(* IEC 61131-3 sources: daoli-st-library/DL_Algo (part 6) *)

(* ---- FC_DL_HumidAirEnthalpy.st ---- *)
(*==============================================================================
 * 组件名称 (Component)  : FC_DL_HumidAirEnthalpy
 * 所属子库 (Sublibrary) : DL_Algo
 * 当前版本 (Version)    : 1.0.1
 * 组件分类 (Category)   : 函数（FUNCTION）· 湿空气热力学算法 · Level 1 算法层
 * 兼容性   (Platform)   : CODESYS 3.5 / TwinCAT 3 / 汇川 InoProShop / Schneider
 *                         Machine Expert；仅依赖 Standard.library（EXP / ABS /
 *                         MIN / MAX），零厂商方言
 * 功能描述 (Function)   : 湿空气比焓 clean-room 计算。公式链：饱和蒸汽压
 *                         p_ws 用 Magnus-Tetens（Stull 参数化，与本库
 *                         FC_DL_DewPointCalc 同系数口径 a=17.625、b=243.04，
 *                         常量复用防两套公式口径漂移）；含湿量
 *                         W = 0.622·phi·p_ws / (p - phi·p_ws)；比焓
 *                         h = 1.006·T + W·(2501 + 1.86·T)。现场用途：洁净
 *                         室/干燥房表冷器与再热功率预算、焓差控制（新风
 *                         焓 < 室内焓 才引入新风）、能耗对比。
 * 出口契约 (Exit)       : 函数返回值 = 湿空气比焓（对应规格引脚表 fEnthalpy
 *                         OUT 列），uErrorId 为 VAR_OUTPUT。异常路径返回
 *                         确定值 0.0，绝不返回未初始化值。
 * 开源溯源 (Origin)     : oscat-building / psychrolib。行为定义对标 OSCAT
 *                         Building 的 AIR_ENTHALPY（0~100 摄氏度域）与
 *                         PsychroLib GetMoistAirEnthalpy 的公开物理公式链；
 *                         公开物理公式无版权义务，不读取、不复制任何源码行，
 *                         100% clean-room 重写并按本库防御规范加严。
 * 属主转移 (R23 裁定)   : Magnus-Tetens 常数（a=17.625、b=243.04）唯一属主
 *                         自 R23 起为 FC_DL_VaporPressureSat；本件内联
 *                         DL_AIR_A / DL_AIR_B 为属主口径的历史引用，本版
 *                         仅声明、逻辑零改动，口径变更以属主件为单一事实源。
 * 规格偏离留档 (R11)    : 规格引脚表 uErrorId 原标注 0001_0203；按第 0 节
 *                         公约 0.7（优先级高于逐组件条款）沿用所在子库
 *                         DL_Algo 既有故障码段 16#0002_xxxx，细分 17xx
 *                         （15xx 露点 / 16xx 流量已占用，顺延无冲突）。
 * 验收向量 (Acceptance) :
 *   V1 T=25.0 RH=60.0 p=101.325：h 约 55.39 kJ/kg 干空气（容差 0.5）；
 *   V2 T=0.0 RH=100.0：h 约 9.44 kJ/kg 干空气（容差 0.5），uErrorId=0；
 *   V3 T=40.0 RH=1.0：干空气端下界，h 约 41.41（容差 0.5）；
 *   V4 RH=0.0：钳位至 1.0，uErrorId=16#0002_1701，照算不发散；
 *   V5 T=150.0：钳位至 100.0，uErrorId=16#0002_1701；
 *   V6 fAtmPress=200.0：钳位至 110.0，uErrorId=16#0002_1702；
 *   V7 T=100.0 RH=100.0：饱和退化分母保护，uErrorId=16#0002_1703，
 *      返回有限确定值；
 *   V8 NaN 输入：拒绝并返回 0.0，uErrorId=16#0002_0004（DL_Algo 公共码）。
 * 故障码表 (Error codes):
 *   16#0002_1701【信息级】温度/湿度越界已钳位照算 / 16#0002_1702【信息级】
 *   大气压越界已钳位照算 / 16#0002_1703【信息级】饱和退化分母已保护 /
 *   16#0002_0004【信息级】输入非有限值已拒绝。全部信息级，本函数无
 *   bError 引脚，故障分级判读经 uErrorId。
 * 修订历史 (Revision)   :
 *   2026-11-15  v1.0.0  首版入库（Round 05 · OSCAT Building 开组 · DL_Algo 补强）
 *============================================================================*)

(*-----------------------------------------------------------------------------
 * 调用示例 (Instance guide)：
 *   fHSupply := FC_DL_HumidAirEnthalpy(fTempC := stAHU.fSupplyT,
 *                                      fRelHum := stAHU.fSupplyRh,
 *                                      uErrorId => uHErr);
 *   fHOutdoor := FC_DL_HumidAirEnthalpy(fTempC := stMet.fTemp,
 *                                       fRelHum := stMet.fRh,
 *                                       fAtmPress := 100.8);
 *   焓差控制联锁：IF (fHOutdoor < fHReturn - 2.0) THEN bFreshAirOk := TRUE;
 *   仅当 uErrorId = 0 时焓值才可用于联锁判断；钳位拍（1701/1702/1703）
 *   的结果按趋势参考处理。
 *----------------------------------------------------------------------------*)

(*-----------------------------------------------------------------------------
 * 常见误用与现场提示 (Field notes)：
 *   1 输入必须是干球温度 + 相对湿度百分数；给成湿球温度或绝对湿度会得到
 *     荒谬结果。露点请先经 FC_DL_DewPointCalc 反算而不是反复试凑本函数。
 *   2 高原/密闭厂房务必传真实大气压 fAtmPress：海拔 2000m 处大气压约
 *     79.5 kPa 已低于钳位下限 80，含湿量 W 会系统性偏小，影响表冷选型。
 *   3 返回值为「每公斤干空气」比焓，做能量平衡时风量要乘干空气密度换算，
 *     勿直接乘湿空气总流量。
 *   4 100 摄氏度/100% 附近 W 发散是物理事实（水的沸点），本函数以 1 Pa
 *     分母下限保护输出有限值，但该域结果无工程意义，勿用于工艺联锁。
 *   5 纯计算无状态，可放心放入高速任务；输入应来自滤波后的温湿度信号。
 *----------------------------------------------------------------------------*)
FUNCTION FC_DL_HumidAirEnthalpy : REAL
VAR_INPUT
    fTempC    : REAL;                    // 干球温度 [摄氏度]，有效域 0.0..100.0 / Dry-bulb temperature [degC], valid range 0.0..100.0
    fRelHum   : REAL;                    // 相对湿度 [百分数]，有效域 1.0..100.0 / Relative humidity [percent], valid range 1.0..100.0
    fAtmPress : REAL := 101.325;         // 大气压 [kPa]，默认标准大气，有效域 80.0..110.0 / Atmospheric pressure [kPa], default standard atmosphere
END_VAR
VAR_OUTPUT
    uErrorId  : UDINT;                   // 故障码，16#0002_0000 = 无故障 / Error code, 16#0002_0000 = no error
END_VAR
VAR
    fTEff     : REAL;                    // 钳位后的生效温度 [摄氏度] / Effective clamped temperature [degC]
    fRhEff    : REAL;                    // 钳位后的生效湿度 [百分数] / Effective clamped humidity [percent]
    fPEff     : REAL;                    // 钳位后的生效大气压 [kPa] / Effective clamped atmospheric pressure [kPa]
    fPws      : REAL;                    // 饱和蒸汽压 [Pa] / Saturation vapor pressure [Pa]
    fPhi      : REAL;                    // 相对湿度份额 [1] / Relative humidity fraction [1]
    fPAbs     : REAL;                    // 绝对大气压 [Pa] / Absolute atmospheric pressure [Pa]
    fPv       : REAL;                    // 水汽分压 [Pa] / Water vapor partial pressure [Pa]
    fDenom    : REAL;                    // 含湿量分母 [Pa] / Humidity ratio denominator [Pa]
    fHumRatio : REAL;                    // 含湿量 [kg 水汽/kg 干空气] / Humidity ratio [kg vapor per kg dry air]
END_VAR
VAR CONSTANT
    DL_AIR_A       : REAL := 17.625;     // Magnus 系数 a [1]，与 FC_DL_DewPointCalc 同口径 / Magnus coefficient a [1], same as dew point FC
    DL_AIR_B       : REAL := 243.04;     // Magnus 系数 b [摄氏度] / Magnus coefficient b [degC]
    DL_AIR_E0      : REAL := 611.2;      // 0 摄氏度饱和水汽压 [Pa] / Saturation vapor pressure at 0 degC [Pa]
    DL_AIR_T_MIN   : REAL := 0.0;        // 温度有效域下限 [摄氏度] / Temperature valid range low [degC]
    DL_AIR_T_MAX   : REAL := 100.0;      // 温度有效域上限 [摄氏度] / Temperature valid range high [degC]
    DL_AIR_RH_MIN  : REAL := 1.0;        // 湿度钳位下限 [百分数]，防 W 比值超线性 / Humidity clamp floor [percent]
    DL_AIR_P_MIN   : REAL := 80.0;       // 大气压钳位下限 [kPa] / Pressure clamp floor [kPa]
    DL_AIR_P_MAX   : REAL := 110.0;      // 大气压钳位上限 [kPa] / Pressure clamp ceiling [kPa]
    DL_AIR_MW      : REAL := 0.622;      // 干空气/水汽摩尔比 [kg/kg] / Molar mass ratio dry air to vapor [kg/kg]
    DL_AIR_CP_DRY  : REAL := 1.006;      // 干空气比热 [kJ/(kg·K)] / Dry air specific heat [kJ/(kg*K)]
    DL_AIR_HFG0    : REAL := 2501.0;     // 0 摄氏度水汽化潜热 [kJ/kg] / Latent heat of vaporization at 0 degC [kJ/kg]
    DL_AIR_CP_VAP  : REAL := 1.86;       // 水汽比热 [kJ/(kg·K)] / Vapor specific heat [kJ/(kg*K)]
    DL_AIR_DENOM_MIN : REAL := 1.0;      // 含湿量分母保护下限 [Pa] / Humidity ratio denominator floor [Pa]
    DL_AIR_EPS     : REAL := 1.0E-6;     // 浮点判零容差 / Float zero tolerance
    DL_AIR_INF_MAX : REAL := 1.0E30;     // 有限值判定幅值上限 / Magnitude bound for finite-value check
END_VAR

(*------------------------------------------------------------------------------
 * 段 1｜出口默认值（IEC 61131-3 强制）：入口即赋确定值，任何提前 RETURN
 *      前输出已确定；异常路径返回 0.0（确定值口径）
 *      Exit defaults (mandatory): outputs assigned deterministically on entry
 *-----------------------------------------------------------------------------*)
FC_DL_HumidAirEnthalpy := 0.0;                    // 返回值（比焓）默认置零 / Return value (enthalpy) preset to zero
uErrorId := 16#0002_0000;                         // 故障码先清零 / Error code cleared first
fTEff := DL_AIR_T_MIN;                            // 温度预置域下限 / Temperature preset to domain floor
fRhEff := DL_AIR_RH_MIN;                          // 湿度预置钳位下限 / Humidity preset to clamp floor
fPEff := 101.325;                                 // 大气压预置标准值 [kPa] / Pressure preset to standard value [kPa]

(*------------------------------------------------------------------------------
 * 段 2｜非有限值防御（公约 0.8）：全部 REAL 输入（含看似常量的大气压）
 *      先做 fX <> fX 检测再比较；命中即拒绝并返回确定值
 *      Non-finite defense: all REAL inputs checked before any comparison
 *-----------------------------------------------------------------------------*)
IF (fTempC <> fTempC) OR (ABS(fTempC) > DL_AIR_INF_MAX)
   OR (fRelHum <> fRelHum) OR (ABS(fRelHum) > DL_AIR_INF_MAX)
   OR (fAtmPress <> fAtmPress) OR (ABS(fAtmPress) > DL_AIR_INF_MAX) THEN
    uErrorId := 16#0002_0004;                     // 输入非有限值已拒绝（DL_Algo 公共码）/ Non-finite input rejected
    FC_DL_HumidAirEnthalpy := 0.0;
    RETURN;
END_IF

(*------------------------------------------------------------------------------
 * 段 3｜温度钳位 [0, 100]：越界信息级码，钳位后照算（R21：不构成故障）
 *      Temperature clamping into [0, 100], info-level code, compute on
 *-----------------------------------------------------------------------------*)
IF (fTempC < DL_AIR_T_MIN) OR (fTempC > DL_AIR_T_MAX) THEN
    fTEff := MIN(MAX(fTempC, DL_AIR_T_MIN), DL_AIR_T_MAX);  // 双侧钳位到有效域 / Two-sided clamp into valid range
    uErrorId := 16#0002_1701;                     // 温度越界已钳位 / Temperature out of range clamped
ELSE
    fTEff := fTempC;                              // 合法温度原值生效 / Valid temperature applied as-is
END_IF

(*------------------------------------------------------------------------------
 * 段 4｜湿度钳位 [1, 100]（公约 0.3 限幅域一致）：下限防 W 发散，上限防
 *      超饱和非物理输入；量纲注释 [百分数] 与限幅域一致（R20）
 *      Humidity clamping into [1, 100], floor guards W divergence
 *-----------------------------------------------------------------------------*)
IF (fRelHum < DL_AIR_RH_MIN) OR (fRelHum > 100.0) THEN
    fRhEff := MIN(MAX(fRelHum, DL_AIR_RH_MIN), 100.0);      // 双侧钳位 / Two-sided clamp
    uErrorId := 16#0002_1701;                     // 湿度越界已钳位 / Humidity out of range clamped
ELSE
    fRhEff := fRelHum;                            // 合法湿度原值生效 / Valid humidity applied as-is
END_IF

(*------------------------------------------------------------------------------
 * 段 5｜大气压钳位 [80, 110] kPa：覆盖海平面 ~ 海拔 2000m 工况域
 *      Atmospheric pressure clamping into [80, 110] kPa
 *-----------------------------------------------------------------------------*)
IF (fAtmPress < DL_AIR_P_MIN) OR (fAtmPress > DL_AIR_P_MAX) THEN
    fPEff := MIN(MAX(fAtmPress, DL_AIR_P_MIN), DL_AIR_P_MAX);  // 双侧钳位 / Two-sided clamp
    uErrorId := 16#0002_1702;                     // 大气压越界已钳位 / Pressure out of range clamped
ELSE
    fPEff := fAtmPress;                           // 合法大气压原值生效 / Valid pressure applied as-is
END_IF

(*------------------------------------------------------------------------------
 * 段 6｜Magnus-Tetens 饱和蒸汽压：与 FC_DL_DewPointCalc 同系数口径，
 *      常量复用防两套公式口径漂移（热平衡算得平）
 *      Magnus-Tetens saturation vapor pressure, same coefficients as dew
 *      point FC, shared constants prevent formula drift
 *-----------------------------------------------------------------------------*)
fPws := DL_AIR_E0 * EXP(DL_AIR_A * fTEff / (DL_AIR_B + fTEff));  // 饱和蒸汽压 [Pa] / Saturation vapor pressure [Pa]

(*------------------------------------------------------------------------------
 * 段 7｜含湿量 W = 0.622·phi·p_ws / (p - phi·p_ws)：分母防除零/防退化
 *      Humidity ratio with denominator guard (divide-by-zero protected)
 *-----------------------------------------------------------------------------*)
fPhi := fRhEff / 100.0;                           // 相对湿度份额 [1] / RH fraction [1]
fPAbs := fPEff * 1000.0;                          // 大气压 kPa → Pa / Pressure kPa converted to Pa
fPv := fPhi * fPws;                               // 水汽分压 [Pa] / Vapor partial pressure [Pa]
fDenom := fPAbs - fPv;                            // 含湿量分母 [Pa] / Denominator [Pa]
IF fPAbs <= DL_AIR_EPS THEN
    uErrorId := 16#0002_1702;                     // 绝对压力退化按大气压类信息级处理 / Degenerate pressure, info code
    FC_DL_HumidAirEnthalpy := 0.0;
    RETURN;
END_IF
IF fDenom <= DL_AIR_DENOM_MIN THEN
    fPv := fPAbs - DL_AIR_DENOM_MIN;              // 饱和退化保护：水汽分压钳至分母下限之上 / Saturation degenerate guard
    uErrorId := 16#0002_1703;                     // 分母退化已保护（100 度/100% 物理发散域） / Degenerate denominator protected
END_IF
fHumRatio := DL_AIR_MW * fPv / (fPAbs - fPv);     // 含湿量 [kg 水汽/kg 干空气] / Humidity ratio [kg/kg dry air]
                                                  // 分母 = fPAbs - fPv ≥ DL_AIR_DENOM_MIN，防除零成立
(*------------------------------------------------------------------------------
 * 段 8｜比焓 h = 1.006·T + W·(2501 + 1.86·T)：显热 + 水汽潜热项
 *      Specific enthalpy: sensible dry-air term plus vapor latent term
 *-----------------------------------------------------------------------------*)
FC_DL_HumidAirEnthalpy := DL_AIR_CP_DRY * fTEff + fHumRatio * (DL_AIR_HFG0 + DL_AIR_CP_VAP * fTEff);
                                                  // 湿空气比焓 [kJ/kg 干空气] / Moist air specific enthalpy [kJ/kg dry air]
END_FUNCTION

(* ---- FC_DL_HystCounterStep.st ---- *)
(*==============================================================================
 * 名称 : FC_DL_HystCounterStep —— 迟滞跨带计数器（上穿 +1 下穿 -1，带位记忆经 nBand 回写）
 * 分类 / 前缀 / 版本 : DL_Algo / FC_DL_ / 1.0.0
 * 溯源 : 开源语义参考（OSCAT/AixOCAT 族，MIT）或 clean-room IEC 实现，未复制源码
 * 平台 : 纯 IEC 61131-3
 * 功能说明 : 以 fUpTh/fDnTh 构成上下带界、fHyst 为校验用回差参考：fIn 上穿
 *            fUpTh 计数 +1，下穿 fDnTh 计数 -1，两界之间不动作（迟滞死区）。
 *            带位记忆 nBand（-1/0/+1）经 VAR_IN_OUT 由调用方持有，保证停在
 *            界外不重复计数、须先穿越对侧门限才反向计数。计数钳位 [nMin,nMax]。
 *            边界处理：fDnTh>=fUpTh、fHyst<0、nMin>nMax 判参数非法；输入
 *            非有限（NaN/±Inf）置 eErr，两种故障下 nBand 保持原值不误动。
 * 错误码 : 16#0001_1C03 = 门限/回差/钳位区间参数非法，或输入非有限（NaN/±Inf）
 *          eErr=0 且 bValid=TRUE 表示计数结果可用（调用方须把返回值写回计数变量）
 * 状态机 : R6 标注 N/A（纯函数无顺序状态，带位记忆由调用方经 nBand 持有，以本节替代 ELSE 兜底）
 * 红线 : R1/R2/R3 ✓ 零全局/零IO/纯IEC ｜ R4 ✓ 非有限拦截/门限校验 ｜ R10 ✓ 标准转换 ｜ R11 ✓ 分号收尾 ｜ R15 ✓ 无保留字撞名
 * 修订记录 : 2026-11-23 v1.0.0 首次入库（R76）
 *============================================================================*)
FUNCTION FC_DL_HystCounterStep : INT
VAR_INPUT
    nCount : INT;      // 当前计数（调用方持有，返回值须写回）/ current count, caller-held
    fIn    : LREAL;    // 被监视输入量 [工程单位] / monitored input value
    fUpTh  : LREAL;    // 上穿计数门限 [工程单位] / up-cross counting threshold
    fDnTh  : LREAL;    // 下穿计数门限 [工程单位] / down-cross counting threshold
    fHyst  : LREAL;    // 回差参考量（须 >=0）[工程单位] / hysteresis reference, must be >= 0
    nMin   : INT;      // 计数下限 [次] / count lower clamp
    nMax   : INT;      // 计数上限 [次] / count upper clamp
END_VAR
VAR_IN_OUT
    nBand  : INT;      // 带位记忆 -1/0/+1（调用方持有回写）/ band memory, caller-held
END_VAR
VAR_OUTPUT
    eErr   : UDINT;    // 故障码，0=正常，1C03=参数非法或非有限 / error code
    bError : BOOL;     // TRUE=本件发生故障 / TRUE when fault occurred
    bValid : BOOL;     // TRUE=计数结果可用 / TRUE when count result is usable
END_VAR
VAR
    _nRet : INT;       // 计数中间值 / count intermediate
END_VAR

FC_DL_HystCounterStep := nCount;             // 返回值预设原计数 / preset return to input count
eErr   := 16#0000_0000;                      // 故障码清零 / clear error code
bError := FALSE;                             // 故障标志清零 / clear error flag
bValid := TRUE;                              // 预设输出可用 / preset valid flag

IF (fIn <> fIn) OR ((fIn - fIn) <> (fIn - fIn))          // fIn 非有限 / NaN or infinite
   OR (fUpTh <> fUpTh) OR ((fUpTh - fUpTh) <> (fUpTh - fUpTh))   // fUpTh 非有限 / NaN or infinite
   OR (fDnTh <> fDnTh) OR ((fDnTh - fDnTh) <> (fDnTh - fDnTh))   // fDnTh 非有限 / NaN or infinite
   OR (fHyst <> fHyst) OR ((fHyst - fHyst) <> (fHyst - fHyst)) THEN  // fHyst 非有限 / NaN or infinite
    eErr   := 16#0001_1C03;                  // 置非有限故障码 / set non-finite code
    bError := TRUE;                          // 置故障标志 / set error flag
    bValid := FALSE;                         // 输出不可用 / outputs not usable
    RETURN;                                  // nBand 冻结原值 / freeze band unchanged
END_IF

IF (fDnTh >= fUpTh) OR (fHyst < 0.0) OR (nMin > nMax) THEN    // 参数合法性校验 / parameter validity check
    eErr   := 16#0001_1C03;                  // 置参数非法码 / set invalid-parameter code
    bError := TRUE;                          // 置故障标志 / set error flag
    bValid := FALSE;                         // 输出不可用 / outputs not usable
    RETURN;                                  // nBand 冻结原值 / freeze band unchanged
END_IF

_nRet := nCount;                             // 取当前计数 / take current count

IF (fIn >= fUpTh) AND (nBand < 1) THEN       // 上穿且非已在高带 / up-cross and not already high
    _nRet := _nRet + 1;                      // 计数 +1 / bump count up
    nBand := 1;                              // 记忆进入高带 / memorize high band
ELSIF (fIn <= fDnTh) AND (nBand > -1) THEN   // 下穿且非已在低带 / down-cross and not already low
    _nRet := _nRet - 1;                      // 计数 -1 / bump count down
    nBand := -1;                             // 记忆进入低带 / memorize low band
ELSIF (fIn > fDnTh) AND (fIn < fUpTh) THEN   // 落入迟滞死区 / inside hysteresis deadband
    nBand := 0;                              // 记忆回到中性带 / memorize neutral band
END_IF

IF _nRet < nMin THEN                         // 计数下限钳位 / clamp lower
    _nRet := nMin;                           // 钳到下限 / clamp to lower
END_IF
IF _nRet > nMax THEN                         // 计数上限钳位 / clamp upper
    _nRet := nMax;                           // 钳到上限 / clamp to upper
END_IF

FC_DL_HystCounterStep := _nRet;              // 回写计数结果 / write back count

END_FUNCTION

(* ---- FC_DL_HystLatchAlarm.st ---- *)
(*==============================================================================
 * 名称 : FC_DL_HystLatchAlarm —— 迟滞触发 + 手动复位锁存报警（状态经 VAR_IN_OUT 由调用方持有）
 * 分类 / 前缀 / 版本 : DL_Algo / FC_DL_ / 1.0.0
 * 溯源 : 开源语义参考（OSCAT/AixOCAT 族，MIT）或 clean-room IEC 实现，未复制源码
 * 平台 : 纯 IEC 61131-3
 * 功能说明 : fIn 上穿 fOn 置位报警并锁存；降到 fOff 以下不自动清除，仅当
 *            bReset=TRUE 才复位（复位后若 fIn 仍 >= fOn 则同拍重新置位，
 *            天然防「复位即复报」盲区）。锁存状态 nState 经 VAR_IN_OUT 由
 *            调用方持有（0=正常 / 1=报警锁存），返回值 = 报警有效电平。
 *            边界处理：fOn<fOff 判参数非法（迟滞反向无意义）；输入非有限
 *            （NaN/±Inf）置 eErr，两种故障下 nState 保持原值不误动。
 * 错误码 : 16#0001_1C02 = 门限次序非法（fOn<fOff），或输入非有限（NaN/±Inf）
 *          eErr=0 且 bValid=TRUE 表示报警电平与 nState 可用
 * 状态机 : R6 标注 N/A（纯函数无顺序状态，锁存态由调用方经 nState 持有，以本节替代 ELSE 兜底）
 * 红线 : R1/R2/R3 ✓ 零全局/零IO/纯IEC ｜ R4 ✓ 非有限拦截/门限校验 ｜ R10 ✓ 标准转换 ｜ R11 ✓ 分号收尾 ｜ R15 ✓ 无保留字撞名
 * 修订记录 : 2026-11-23 v1.0.0 首次入库（R76）
 *============================================================================*)
FUNCTION FC_DL_HystLatchAlarm : BOOL
VAR_INPUT
    fIn    : LREAL;    // 被监视输入量 [工程单位] / monitored input value
    fOn    : LREAL;    // 报警置位门限 [工程单位] / alarm set threshold
    fOff   : LREAL;    // 迟滞参考门限（仅作参数校验：要求 fOn >= fOff）[工程单位] / hysteresis reference, param check only
    bReset : BOOL;     // 复位指令（沿/电平均可，调用方决定）/ reset command
END_VAR
VAR_IN_OUT
    nState : INT;      // 锁存状态 0=正常 1=报警（调用方持有回写）/ latched state, caller-held
END_VAR
VAR_OUTPUT
    eErr   : UDINT;    // 故障码，0=正常，1C02=参数非法或非有限 / error code
    bError : BOOL;     // TRUE=本件发生故障 / TRUE when fault occurred
    bValid : BOOL;     // TRUE=报警电平可用 / TRUE when alarm level is usable
END_VAR

FC_DL_HystLatchAlarm := FALSE;               // 报警电平预设 FALSE / preset alarm to FALSE
eErr   := 16#0000_0000;                      // 故障码清零 / clear error code
bError := FALSE;                             // 故障标志清零 / clear error flag
bValid := TRUE;                              // 预设输出可用 / preset valid flag

IF (fIn <> fIn) OR ((fIn - fIn) <> (fIn - fIn))          // fIn 非有限 / NaN or infinite
   OR (fOn <> fOn) OR ((fOn - fOn) <> (fOn - fOn))        // fOn 非有限 / NaN or infinite
   OR (fOff <> fOff) OR ((fOff - fOff) <> (fOff - fOff)) THEN  // fOff 非有限 / NaN or infinite
    eErr   := 16#0001_1C02;                  // 置非有限故障码 / set non-finite code
    bError := TRUE;                          // 置故障标志 / set error flag
    bValid := FALSE;                         // 输出不可用 / outputs not usable
    RETURN;                                  // nState 冻结原值，不误动 / freeze state unchanged
END_IF

IF fOn < fOff THEN                           // 迟滞反向：参数非法 / reversed hysteresis invalid
    eErr   := 16#0001_1C02;                  // 置参数非法码 / set invalid-parameter code
    bError := TRUE;                          // 置故障标志 / set error flag
    bValid := FALSE;                         // 输出不可用 / outputs not usable
    RETURN;                                  // nState 冻结原值 / freeze state unchanged
END_IF

IF bReset THEN                               // 手动复位优先（先清后判）/ reset first, judge after
    nState := 0;                             // 清除锁存 / clear latch
END_IF
IF nState = 0 THEN                           // 非锁存态才可置位 / only unlatched state can set
    IF fIn >= fOn THEN                       // 上穿置位门限 / rising past set threshold
        nState := 1;                         // 置位并锁存 / set and latch
    END_IF
END_IF

FC_DL_HystLatchAlarm := (nState = 1);        // 回写报警电平 / write back alarm level

END_FUNCTION

(* ---- FC_DL_HystTimeQualified.st ---- *)
(*==============================================================================
 * 名称 : FC_DL_HystTimeQualified —— 迟滞 + 时间确认翻转（确认计时由调用方 TON 持有）
 * 分类 / 前缀 / 版本 : DL_Algo / FC_DL_ / 1.0.0
 * 溯源 : 开源语义参考（OSCAT/AixOCAT 族，MIT）或 clean-room IEC 实现，未复制源码
 * 平台 : 纯 IEC 61131-3
 * 功能说明 : 输出翻转需时间确认：bRawIn=FALSE 时输出立即 FALSE 且确认计时
 *            清零（tNewElapsed=T#0s）；bRawIn=TRUE 且输出当前 FALSE 时，仅当
 *            调用方 TON 累计 tElapsed >= tQual 才翻转 TRUE；输出已 TRUE 且
 *            原始输入仍 TRUE 则保持。tElapsed 语义 = 调用方 TON.ET（bRawIn
 *            期间单调增长），tNewElapsed 回传给调用方供下一拍使用。
 *            边界处理：tQual<=T#0s 视为立即确认（0 时延合法用法）；
 *            bPrevOut=TRUE 而 bRawIn=FALSE 时立即翻 FALSE（OFF 无延时）。
 * 错误码 : 16#0001_1C04 为本件预留码位（当前实现无故障路径），eErr 恒 0、bValid 恒 TRUE
 * 状态机 : R6 标注 N/A（纯函数无顺序状态，确认计时由调用方 TON 持有，以本节替代 ELSE 兜底）
 * 红线 : R1/R2/R3 ✓ 零全局/零IO/纯IEC ｜ R4 ✓ 时间比较口径明确 ｜ R10 ✓ 标准转换 ｜ R11 ✓ 分号收尾 ｜ R15 ✓ 无保留字撞名
 * 修订记录 : 2026-11-23 v1.0.0 首次入库（R76）
 *============================================================================*)
FUNCTION FC_DL_HystTimeQualified : BOOL
VAR_INPUT
    bRawIn   : BOOL;   // 原始输入（未经确认）/ raw input before qualification
    tQual    : TIME;   // 确认时长门限 [ms] / qualification duration threshold
    bPrevOut : BOOL;   // 上一拍输出（调用方持有）/ previous output, caller-held
    tElapsed : TIME;   // 调用方 TON 累计确认时间 [ms] / caller-held TON elapsed time
END_VAR
VAR_OUTPUT
    tNewElapsed : TIME;    // 回传确认时间（供调用方下一拍使用）/ elapsed time passed back to caller
    eErr        : UDINT;   // 故障码，0=正常（本件无故障路径）/ error code, 0=ok (no fault path)
    bError      : BOOL;    // 故障标志，恒 FALSE / error flag, always FALSE
    bValid      : BOOL;    // TRUE=输出与计时可用，恒 TRUE / TRUE when outputs are usable
END_VAR

eErr        := 16#0000_0000;             // 故障码清零 / clear error code
bError      := FALSE;                    // 故障标志清零 / clear error flag
bValid      := TRUE;                     // 本件无故障路径，恒可用 / always valid
tNewElapsed := T#0s;                     // 确认计时预设清零 / preset elapsed to zero

IF NOT bRawIn THEN                       // 原始输入失效：OFF 无延时 / raw input low: immediate off
    FC_DL_HystTimeQualified := FALSE;    // 输出立即 FALSE / output FALSE immediately
    tNewElapsed := T#0s;                 // 确认计时清零（调用方应同步复位 TON）/ reset qualification timer
    RETURN;                              // 提前收口 / early exit
END_IF

tNewElapsed := tElapsed;                 // 原始输入有效：计时透传 / raw high: pass timer through

IF bPrevOut THEN                         // 输出已 TRUE 且原始输入仍 TRUE / already on and raw high
    FC_DL_HystTimeQualified := TRUE;     // 保持 TRUE / keep TRUE
ELSIF tElapsed >= tQual THEN             // 确认计时到限 / qualification time reached
    FC_DL_HystTimeQualified := TRUE;     // 翻转为 TRUE / flip to TRUE
ELSE                                     // 确认时间未到 / qualification not reached
    FC_DL_HystTimeQualified := FALSE;    // 维持 FALSE / keep FALSE
END_IF

END_FUNCTION

(* ---- FC_DL_HystWindow3.st ---- *)
(*==============================================================================
 * 名称 : FC_DL_HystWindow3 —— 三带迟滞带位判定（低/中/高，回差记忆由调用方持有）
 * 分类 / 前缀 / 版本 : DL_Algo / FC_DL_ / 1.0.0
 * 溯源 : 开源语义参考（OSCAT/AixOCAT 族，MIT）或 clean-room IEC 实现，未复制源码
 * 平台 : 纯 IEC 61131-3
 * 功能说明 : 返回三带带位：0=低带、1=中带、2=高带。上行走「上行门限」进带
 *            （fIn>=fLowOn 进中带、fIn>=fHighOn 进高带），下行走「下行门限」
 *            退带（fIn<fLowOff 退低带、fIn<fHighOff 退中带），回差由门限对
 *            (fLowOn/fLowOff) 与 (fHighOn/fHighOff) 构成，历史带位经
 *            nPrevState 由调用方持有回传。
 *            边界处理：fLowOff<=fLowOn<fHighOff<=fHighOn 不满足判参数非法
 *            （eErr、返回 0、bValid=FALSE）；nPrevState 非 0/1/2 时走 ELSE
 *            兜底按电平重判；输入非有限（NaN/±Inf）置 eErr。
 * 错误码 : 16#0001_1C01 = 门限次序非法（不满足 fLowOff<=fLowOn<fHighOff<=fHighOn），或输入非有限
 *          eErr=0 且 bValid=TRUE 表示带位可用
 * 状态机 : R6 标注 N/A（纯函数无顺序状态，带位记忆由调用方持有，本件以 ELSE 兜底替代 CASE 收口）
 * 红线 : R1/R2/R3 ✓ 零全局/零IO/纯IEC ｜ R4 ✓ 非有限拦截/门限校验 ｜ R10 ✓ 标准转换 ｜ R11 ✓ 分号收尾 ｜ R15 ✓ 无保留字撞名
 * 修订记录 : 2026-11-23 v1.0.0 首次入库（R76）
 *============================================================================*)
FUNCTION FC_DL_HystWindow3 : INT
VAR_INPUT
    fIn       : LREAL;   // 被判定输入量 [工程单位] / input value under test
    fLowOn    : LREAL;   // 低带→中带上行门限 [工程单位] / rising threshold low-to-mid
    fLowOff   : LREAL;   // 中带→低带下行门限 [工程单位] / falling threshold mid-to-low
    fHighOn   : LREAL;   // 中带→高带上行门限 [工程单位] / rising threshold mid-to-high
    fHighOff  : LREAL;   // 高带→中带下行门限 [工程单位] / falling threshold high-to-mid
    nPrevState: INT;     // 上一拍带位 0/1/2（调用方持有）/ previous band, caller-held
END_VAR
VAR_OUTPUT
    eErr   : UDINT;    // 故障码，0=正常，1C01=参数非法或非有限 / error code
    bError : BOOL;     // TRUE=本件发生故障 / TRUE when fault occurred
    bValid : BOOL;     // TRUE=带位可用 / TRUE when band is usable
END_VAR
VAR
    _nRet : INT;       // 带位计算中间值 / band intermediate
END_VAR

FC_DL_HystWindow3 := 0;                      // 带位预设 0（低带）/ preset band to low
eErr   := 16#0000_0000;                      // 故障码清零 / clear error code
bError := FALSE;                             // 故障标志清零 / clear error flag
bValid := TRUE;                              // 预设输出可用 / preset valid flag

IF (fIn <> fIn) OR ((fIn - fIn) <> (fIn - fIn))            // fIn 非有限 / NaN or infinite
   OR (fLowOn <> fLowOn) OR ((fLowOn - fLowOn) <> (fLowOn - fLowOn))   // fLowOn 非有限 / NaN or infinite
   OR (fLowOff <> fLowOff) OR ((fLowOff - fLowOff) <> (fLowOff - fLowOff)) // fLowOff 非有限 / NaN or infinite
   OR (fHighOn <> fHighOn) OR ((fHighOn - fHighOn) <> (fHighOn - fHighOn)) // fHighOn 非有限 / NaN or infinite
   OR (fHighOff <> fHighOff) OR ((fHighOff - fHighOff) <> (fHighOff - fHighOff)) THEN  // fHighOff 非有限 / NaN or infinite
    eErr   := 16#0001_1C01;                  // 置非有限故障码 / set non-finite code
    bError := TRUE;                          // 置故障标志 / set error flag
    bValid := FALSE;                         // 带位不可用 / band not usable
    RETURN;                                  // 返回 0 / return zero
END_IF

IF NOT ((fLowOff <= fLowOn) AND (fLowOn < fHighOff) AND (fHighOff <= fHighOn)) THEN    // 门限次序校验 / threshold order check
    eErr   := 16#0001_1C01;                  // 置参数非法码 / set invalid-parameter code
    bError := TRUE;                          // 置故障标志 / set error flag
    bValid := FALSE;                         // 带位不可用 / band not usable
    RETURN;                                  // 返回 0 / return zero
END_IF

_nRet := nPrevState;                         // 取上一拍带位 / take previous band

IF _nRet = 0 THEN                            // 低带滞回分支 / low band hysteresis branch
    IF fIn >= fLowOn THEN                    // 上穿中带门限 / rising past mid entry
        _nRet := 1;                          // 进中带 / enter mid band
    END_IF
ELSIF _nRet = 1 THEN                         // 中带滞回分支 / mid band hysteresis branch
    IF fIn >= fHighOn THEN                   // 上穿高带门限 / rising past high entry
        _nRet := 2;                          // 进高带 / enter high band
    ELSIF fIn < fLowOff THEN                 // 下穿低带退出门限 / falling past low exit
        _nRet := 0;                          // 退低带 / fall to low band
    END_IF
ELSIF _nRet = 2 THEN                         // 高带滞回分支 / high band hysteresis branch
    IF fIn < fHighOff THEN                   // 下穿中带退出门限 / falling past mid exit
        _nRet := 1;                          // 退中带 / fall to mid band
    END_IF
ELSE                                         // ELSE 兜底：非法带位按电平重判 / else: re-judge by level
    IF fIn >= fHighOn THEN                   // 电平在高带门限上 / level above high entry
        _nRet := 2;                          // 判高带 / judge high band
    ELSIF fIn >= fLowOn THEN                 // 电平在中带门限上 / level above low entry
        _nRet := 1;                          // 判中带 / judge mid band
    ELSE                                     // 电平在低带 / level in low band
        _nRet := 0;                          // 判低带 / judge low band
    END_IF
END_IF

FC_DL_HystWindow3 := _nRet;                  // 回写带位 / write back band

END_FUNCTION

(* ---- FC_DL_IllinoisIterStep.st ---- *)
(* ============================================================
   DL_Algo / FC_DL_IllinoisIterStep ｜ v1.0.0 ｜ 2026-11-25
   功能：Illinois 改进试位单步的端点修正环节。由上次插值点 fXPrev 落在括号哪一半
         定出本次替换侧（1=a / 2=b）；若与 uLastSide 相同（同端连续被保留），
         则把停滞端函数值折半，防单侧卡死（收敛阶高于经典试位法）
   边界：端点函数值判零（容差）→ 已是根，不折半原样回传；非有限 → 两值写 0
         且 uSideOut=0（上层据侧码 0 拒收本步，N1：判据位与实值同源）
   依赖：仅 IEC 61131-3（ABS / MIN / MAX） ｜ 溯源：DLF-B-ROOTSTEP（内部原创线）
   ============================================================ *)
FUNCTION FC_DL_IllinoisIterStep : BOOL
VAR_INPUT
    fA        : LREAL;  // 括号下界 [-] / Lower bracket bound
    fB        : LREAL;  // 括号上界 [-] / Upper bracket bound
    fFa       : LREAL;  // 下界函数值 [-] / Function value at the lower bound
    fFb       : LREAL;  // 上界函数值 [-] / Function value at the upper bound
    fXPrev    : LREAL;  // 上次弦线插值点 [-] / Previous interpolated point
    uLastSide : UDINT;  // 上次被替换侧 0 无历史 / 1 a / 2 b [-] / Side replaced last time
END_VAR
VAR_OUTPUT
    fFaOut       : LREAL;  // a 端函数值（可能折半）[-] / Outgoing value at the lower bound
    fFbOut       : LREAL;  // b 端函数值（可能折半）[-] / Outgoing value at the upper bound
    uSideOut     : UDINT;  // 本次替换侧 0 非法 / 1 a / 2 b [-] / Side replaced this time
    bHalfApplied : BOOL;   // 本次执行了停滞端折半 [-] / Stagnating endpoint halving applied
END_VAR
VAR
    _fMid  : LREAL;  // 括号中点 [-] / Bracket midpoint
    _uSide : UDINT;  // 本次替换侧暂存 [-] / Staged side code
END_VAR
VAR CONSTANT
    DL_ILL_EPS : LREAL := 1.0E-12;  // 判零容差 [-] / Zero tolerance
END_VAR

(* 段 0：出口预置（侧码 0、未折半，值域先落 0） *)
FC_DL_IllinoisIterStep := FALSE;
fFaOut := 0.0;  fFbOut := 0.0;  uSideOut := 0;  bHalfApplied := FALSE;

(* 段 1：非有限闸（NaN 自反 + Inf 差值自减，五入参全量枚举，R79/R272） *)
IF (fA <> fA) OR (fB <> fB) OR (fFa <> fFa) OR (fFb <> fFb) OR (fXPrev <> fXPrev) THEN
    RETURN;
END_IF
(* Inf 双判须覆盖 fA/fB/fFa/fFb：只判 fXPrev 时 fFa=+Inf 会原样进 fFaOut 出口并
   以 uSideOut≠0、返回 TRUE 上报（伪有效端点值） *)
IF ((fA - fA) <> (fA - fA)) OR ((fB - fB) <> (fB - fB))
   OR ((fFa - fFa) <> (fFa - fFa)) OR ((fFb - fFb) <> (fFb - fFb))
   OR ((fXPrev - fXPrev) <> (fXPrev - fXPrev)) THEN RETURN; END_IF
fFaOut := fFa;  fFbOut := fFb;                // 闸后先原样回传

(* 段 2：端点已是根（容差判零）则不做任何修正 *)
IF (ABS(fFa) <= DL_ILL_EPS) OR (ABS(fFb) <= DL_ILL_EPS) THEN
    uSideOut := 1;  FC_DL_IllinoisIterStep := TRUE;  RETURN;
END_IF

(* 段 3：本次替换侧判定（上次插值点落在哪一半） *)
_fMid := MIN(fA, fB) + (ABS(fB - fA)) / 2.0;
IF fXPrev <= _fMid THEN
    _uSide := 1;                              // 偏下：a 端被替换
ELSE
    _uSide := 2;                              // 偏上：b 端被替换
END_IF

(* 段 4：Illinois 折半规则（同一端连续被保留 → 停滞端折半） *)
IF uLastSide = _uSide THEN
    IF _uSide = 1 THEN
        fFbOut := fFb / 2.0;                  // a 被替换：停滞端为 b
    ELSE
        fFaOut := fFa / 2.0;                  // b 被替换：停滞端为 a
    END_IF
    bHalfApplied := TRUE;
END_IF

(* 段 5：单一出口裁决（N4） *)
uSideOut := _uSide;  FC_DL_IllinoisIterStep := TRUE;
END_FUNCTION

(* ---- FC_DL_IterTermJudge.st ---- *)
(* ============================================================
   DL_Algo / FC_DL_IterTermJudge ｜ v1.0.0 ｜ 2026-11-25
   功能：迭代终止四判据仲裁，优先级 超时 > 迭代上限 > 区间宽度 > 步长；
         命中即 bDone=TRUE 并给 uReason：0 继续 / 1 宽度 / 2 步长 / 3 上限 / 4 超时
   边界：容差与超时按 R95 代理阈值三句声明 —— 代理值：宽度 1E-9、步长 1E-9、
         超时 10s；覆盖 1~100ms 常规控制周期；覆盖不到的亚毫秒任务与超长批处理
         由调用方自备阈值件负责。5 号码反证：NaN 输入下四判据比较全假 → 永不终止，
         该死锁无法由 0~4 号组合观测，故立 5 号（R90）
   依赖：仅 IEC 61131-3（ABS / TIME_TO_REAL） ｜ 溯源：DLF-B-ROOTSTEP（内部原创线）
   ============================================================ *)
FUNCTION FC_DL_IterTermJudge : BOOL
VAR_INPUT
    fWidth   : LREAL;  // 当前括号宽度，域 ≥ 0 [-] / Current bracket width
    fStep    : LREAL;  // 上一步位移绝对值，域 ≥ 0 [-] / Absolute step of the last iteration
    uIter    : UDINT;  // 已用迭代次数 [次] / Iterations already consumed
    uIterMax : UDINT;  // 允许最大迭代次数，0 = 不限 [次] / Iteration cap, zero means unlimited
    tElapsed : TIME;   // 已耗时 [ms] / Elapsed time since the iteration started
END_VAR
VAR_OUTPUT
    bDone   : BOOL;   // 终止标志 [-] / Terminate flag
    uReason : UDINT;  // 终止原因码 0/1/2/3/4/5 [-] / Termination reason code
END_VAR
VAR
    _fTEsc : LREAL;  // 超时阈值秒值 [s] / Timeout threshold in seconds
    _fElap : LREAL;  // 已耗时秒值 [s] / Elapsed time in seconds
END_VAR
VAR CONSTANT
    DL_ITJ_XTOL : LREAL := 1.0E-9;  // 区间宽度容差代理值 [-] / Proxy tolerance on the bracket width
    DL_ITJ_STOL : LREAL := 1.0E-9;  // 步长容差代理值 [-] / Proxy tolerance on the step size
    DL_ITJ_TMAX : TIME := T#10S;    // 超时阈值代理值 [ms] / Proxy timeout value
    DL_ITJ_MSPS : LREAL := 1000.0;  // 毫秒 → 秒换算系数 [ms/s] / Milliseconds per second
END_VAR

(* 段 0：出口预置安全侧（不终止、原因 0） *)
FC_DL_IterTermJudge := FALSE;
bDone := FALSE;  uReason := 0;

(* 段 1：非有限闸（判据量不可用 → 安全侧终止，防死锁） *)
IF (fWidth <> fWidth) OR (fStep <> fStep)
   OR ((fWidth - fWidth) <> (fWidth - fWidth)) OR ((fStep - fStep) <> (fStep - fStep)) THEN
    bDone := TRUE;  uReason := 5;  RETURN;
END_IF

(* 段 2：超时判据（最高优先级，时间域不可回退） *)
_fTEsc := TIME_TO_REAL(DL_ITJ_TMAX) / DL_ITJ_MSPS;
_fElap := TIME_TO_REAL(tElapsed) / DL_ITJ_MSPS;
IF _fElap >= _fTEsc THEN bDone := TRUE;  uReason := 4;  RETURN; END_IF

(* 段 3：迭代上限判据（uIterMax = 0 视为不限） *)
IF (uIterMax > 0) AND (uIter >= uIterMax) THEN bDone := TRUE;  uReason := 3;  RETURN; END_IF

(* 段 4：区间宽度判据 *)
IF ABS(fWidth) <= DL_ITJ_XTOL THEN bDone := TRUE;  uReason := 1;  RETURN; END_IF

(* 段 5：步长判据（最后一级，防「步长极小但区间仍宽」的假收敛） *)
IF ABS(fStep) <= DL_ITJ_STOL THEN bDone := TRUE;  uReason := 2;  RETURN; END_IF

(* 段 6：单一出口裁决（N4：未命中任何判据才继续） *)
bDone := FALSE;  uReason := 0;  FC_DL_IterTermJudge := TRUE;
END_FUNCTION

(* ---- FC_DL_Median3Vote.st ---- *)
// FC_DL_Median3Vote v1.0.0
(*==============================================================================
 * 功能描述: 三取二中值表决。三输入排序取中值输出；极差 (max-min) 超 fSpreadThr
 *           置 bSpread 诊断（输入分歧大，表决可信度降级）；任一输入非有限 →
 *           bValid=FALSE 并返回 0。
 * 接口契约: 输入 fA/fB/fC/fSpreadThr；输出 bValid/bSpread，返回中值。
 * 修订历史: 2026-11-23  v1.0.0  R74 首版
 *==============================================================================*)

FUNCTION FC_DL_Median3Vote : REAL
VAR_INPUT
    fA         : REAL := 0.0;   // 表决输入 A [工程单位] / Vote input A
    fB         : REAL := 0.0;   // 表决输入 B [工程单位] / Vote input B
    fC         : REAL := 0.0;   // 表决输入 C [工程单位] / Vote input C
    fSpreadThr : REAL := 1.0;   // 极差诊断阈值，域 > 0 [工程单位] / Spread diagnosis threshold
END_VAR
VAR_OUTPUT
    bValid  : BOOL;             // 结果有效回执 [-] / Result validity receipt
    bSpread : BOOL;             // 极差超阈诊断标志 [-] / Spread over threshold flag
END_VAR
VAR
    fMax : REAL;                // 三输入最大值 [工程单位] / Maximum of the three
    fMin : REAL;                // 三输入最小值 [工程单位] / Minimum of the three
END_VAR

(* —— 段 0：全路径赋值缺省（无效安全侧） —— *)
bValid := FALSE;                             // 有效回执预清 / Validity preset
bSpread := FALSE;                            // 分歧诊断预清 / Spread preset
FC_DL_Median3Vote := 0.0;                    // 返回值缺省零 / Result default zero

(* —— 段 1：非有限闸（任一 NaN 即表决失效） —— *)
IF (fA <> fA) OR (fB <> fB) OR (fC <> fC) THEN   // NaN 自反判（判等禁令唯一例外） / NaN self-reflexive tests
    RETURN;                                  // 无效返回零 / Invalid, return zero
END_IF

(* —— 段 2：极值派生与中值合成（中值 = 和 - 最大 - 最小，三值和幅值受输入域约束） —— *)
fMax := MAX(MAX(fA, fB), fC);                // 三输入最大值 / Maximum of the three
fMin := MIN(MIN(fA, fB), fC);                // 三输入最小值 / Minimum of the three
IF ABS(fMax) >= 1.0E38 THEN                  // 近 Inf 幅值闸 / Near-Inf magnitude gate
    RETURN;                                  // 无效返回零 / Invalid, return zero
END_IF
FC_DL_Median3Vote := (fA + fB + fC) - fMax - fMin;   // 中值合成（三值代数恒等式） / Median by algebraic identity
bValid := TRUE;                              // 有效回执 / Validity receipt
IF fSpreadThr > 0.0 THEN                     // 阈值正值闸（R4 防无效比较域） / Threshold positive gate
    bSpread := (fMax - fMin) > fSpreadThr;   // 极差超阈诊断 / Spread over threshold diagnosis
END_IF

END_FUNCTION

(* ---- FC_DL_MixAirStateCalc.st ---- *)
//==============================================================================
// 函数：FC_DL_MixAirStateCalc ｜ 中文名称：回风/新风混合点状态计算（焓湿图族拆分⑤）
// 所属子库：DL_Algo ｜ 版本：v1.0.2 ｜ 兼容：CODESYS V3.5+ / TwinCAT 3 / 汇川 InoProShop
// 功能描述：质量守恒加权求回风/新风混合点状态：干球温度与含湿量分别按
//           新风比加权（fMixX = fOaFrac/100·fOaX + (1−fOaFrac/100)·fRaX），
//           并内联复算混合焓 h = 1.006·T + W·(2501 + 1.86·T) [kJ/kg 干空气]；
//           结露判据用混合点水汽分压与混合温度下饱和压比较（p_v_mix >
//           p_ws(T_mix) 即越过饱和线），饱和压取自族属主
//           FC_DL_VaporPressureSat，零内联公式。ASHRAE 混风质量守恒公开
//           公式；职责边界：本件算状态点，经济器决策属 FB_DL_EnthalpyCompareCtrl。
// 开源溯源 (Origin)：改写自 OSCAT Building 行为定义（OSCAT 许可，仅行为定义，零代码行）——道莅 clean-room 实现
// 单位表：T[°C] / W[kg 水蒸气/kg 干空气] / 新风比[%] / h[kJ/kg 干空气] /
//         p[Pa] / p_v[Pa] / p_ws[Pa]
// 错误码表：16#0002_3101 信息级（新风比或含湿量域外已钳位，不置 bError）/
//           16#0002_3110 故障级（任一输入非有限，置 bError）/
//           16#0002_3102、16#0002_3111、16#0002_3112 预留禁用（不得挪用）
// 状态机：N/A（纯函数，无状态）
// 边界行为：① fOaFrac 域外（0~100 外）→ 钳位 + 信息 3101；② 任一输入
//           非有限 → 故障 3110、bValid := FALSE、输出 0；③ 含湿量输入
//           < 0 → 钳 0 + 信息 3101 复用（R90）；④ 结露仅置 bCondensation
//           预警位，不置故障（结露是工况事实不是错误）；⑤ 属主件拒绝 →
//           故障 3110 复用（R90）；异常路径输出确定值，绝不输出未初始化值。
// 依赖收窄 (R11 留档③)：DL_Algo 不得跨库调用，混合焓用本件内联等价式
//           h := 1.006·T + W·(2501 + 1.86·T)，与 FC_DL_HumidAirEnthalpy 的
//           口径一致性由本件头注释承担验证责任（常量逐一同源：1.006 /
//           2501 / 1.86，改动任一侧须同步复核另一侧）。
// 修订历史：v1.0.0 2026-11-17 首版（R23 派单 · T1-2 焓湿图族拆分⑤ · 族收口件）
//           v1.0.1 2026-11-17 R23 终审修复：段 2 非有限闸补查 fOaFrac
//           （原漏判 NaN 新风比会以 bValid=TRUE 放行 NaN 混合输出），契约不变。
//           v1.0.2 2026-11-23 R73 补 bValid 回执：段 6 属主件调用补收 bValid
//           局部回执，回执无效并入既有 3110 兜底分支，契约不变。
//==============================================================================

(*------------------------------------------------------------------------------
 * 调用示例：bOk := FC_DL_MixAirStateCalc(
 *             fRaTempC := 26.0, fRaHumRatio := 0.0105,
 *             fOaTempC := 33.0, fOaHumRatio := 0.0192,
 *             fOaFrac := 30.0, fPress := 101325.0,
 *             fMixTempC => fTmix, fMixHumRatio => fWmix,
 *             fMixEnthalpy => fHmix, bCondensation => bCond, eErr => uE);
 * 结露预警口径：bCondensation = TRUE 时混合点位于饱和线下游，表冷器/风道
 * 有凝水风险；该位是工况事实，上层据此决策，不作为故障联锁。
 *-----------------------------------------------------------------------------*)
FUNCTION FC_DL_MixAirStateCalc : BOOL
VAR_INPUT
    fRaTempC     : LREAL;                  // 回风干球温度 [摄氏度] / Return-air dry-bulb temperature [degC]
    fRaHumRatio  : LREAL;                  // 回风含湿量 [kg 水蒸气/kg 干空气] / Return-air humidity ratio [kg/kg dry air]
    fOaTempC     : LREAL;                  // 新风干球温度 [摄氏度] / Outdoor-air dry-bulb temperature [degC]
    fOaHumRatio  : LREAL;                  // 新风含湿量 [kg 水蒸气/kg 干空气] / Outdoor-air humidity ratio [kg/kg dry air]
    fOaFrac      : LREAL;                  // 新风比 [百分数]，有效域 0.0..100.0，域外钳位照算 / Outdoor-air fraction [percent], valid range 0.0..100.0
    fPress       : LREAL := 101325.0;      // 大气压 [Pa]，引脚注入非魔法数 / Atmospheric pressure [Pa], injected via the pin
END_VAR
VAR_OUTPUT
    fMixTempC    : LREAL;                  // 混合点干球温度 [摄氏度] / Mixed dry-bulb temperature [degC]
    fMixHumRatio : LREAL;                  // 混合点含湿量 [kg 水蒸气/kg 干空气] / Mixed humidity ratio [kg/kg dry air]
    fMixEnthalpy : LREAL;                  // 混合点比焓 [kJ/kg 干空气] / Mixed specific enthalpy [kJ/kg dry air]
    bCondensation: BOOL;                   // TRUE = 混合点越过饱和线，结露预警（非故障） / TRUE = mixing point crosses the saturation line, condensation warning, not a fault
    eErr         : UDINT;                  // 错误码，0 = 无错 / Error code, 0 = no error
    bError       : BOOL;                   // 故障级标志，仅故障级错误置位 / Fault-class flag, set only on fault-level codes
    bValid       : BOOL;                   // 输出可用标志 / Outputs usable flag
END_VAR
VAR CONSTANT
    DL_MIX_CP_DRY  : LREAL := 1.006;     // 干空气比热 [kJ/(kg·K)]，与 FC_DL_HumidAirEnthalpy 同源 / Dry-air specific heat [kJ/(kg*K)], same source as the enthalpy FC
    DL_MIX_HFG0    : LREAL := 2501.0;    // 0 摄氏度水汽化潜热 [kJ/kg]，同源口径 / Latent heat of vaporization at 0 degC [kJ/kg], same source
    DL_MIX_CP_VAP  : LREAL := 1.86;      // 水汽比热 [kJ/(kg·K)]，同源口径 / Vapor specific heat [kJ/(kg*K)], same source
    DL_MIX_MW      : LREAL := 0.621945;  // 干空气/水蒸气摩尔质量比 [kg/kg]，ASHRAE 口径 / Molar mass ratio dry air to vapor [kg/kg], ASHRAE
    DL_MIX_FRAC_MIN: LREAL := 0.0;       // 新风比钳位下限 [百分数] / Outdoor fraction clamp floor [percent]
    DL_MIX_FRAC_MAX: LREAL := 100.0;     // 新风比钳位上限 [百分数] / Outdoor fraction clamp ceiling [percent]
    DL_MIX_EPS     : LREAL := 1.0E-6;    // 浮点判零容差 [Pa] / Float zero tolerance [Pa]
    DL_MIX_INF     : LREAL := 1.7976931348623157E308; // LREAL 幅值上限 / LREAL magnitude ceiling
END_VAR
VAR
    fFracEff   : LREAL;                  // 钳位后的生效新风比份额 [1] / Effective outdoor fraction share [1]
    fRaWEff    : LREAL;                  // 钳位后的生效回风含湿量 [kg/kg] / Effective return-air humidity ratio [kg/kg]
    fOaWEff    : LREAL;                  // 钳位后的生效新风含湿量 [kg/kg] / Effective outdoor-air humidity ratio [kg/kg]
    fPvMix     : LREAL;                  // 混合点水汽分压 [Pa] / Mixed vapor partial pressure [Pa]
    fPwsMix    : LREAL;                  // 混合温度下饱和压 [Pa]，属主件取得 / Saturation pressure at the mixed temperature [Pa]
    fDenom     : LREAL;                  // 分压反算分母 (MW + W_mix) [kg/kg] / Denominator of the partial-pressure inversion [kg/kg]
    _bPwsValid : BOOL;                   // 饱和压属主件输出可用回执 / Saturation owner FC outputs-usable receipt
    _bPwsClamped : BOOL;    // 属主件钳位回执（本件不消费，仅契约全回执） / Owner clamp receipt (unused, full-receipt contract)
    _nPwsErr     : UDINT;   // 属主件错误码回执 / Owner error-code receipt
    _bPwsError   : BOOL;    // 属主件故障级回执 / Owner fault-flag receipt
END_VAR

(*------------------------------------------------------------------------------
 * 段 1｜出口默认值：入口即赋确定值
 *      Exit defaults: outputs assigned deterministically on entry
 *-----------------------------------------------------------------------------*)
FC_DL_MixAirStateCalc := FALSE;          // 返回值默认无效 / Return value preset invalid
fMixTempC := 0.0;                        // 混合温度默认置零 / Mixed temperature preset to zero
fMixHumRatio := 0.0;                     // 混合含湿量默认置零 / Mixed humidity ratio preset to zero
fMixEnthalpy := 0.0;                     // 混合焓默认置零 / Mixed enthalpy preset to zero
bCondensation := FALSE;                  // 结露预警默认 FALSE / Condensation warning preset FALSE
eErr := 16#0000_0000;                    // 错误码先清零 / Error code cleared first
bError := FALSE;                         // 故障标志先清零 / Fault flag cleared first
bValid := FALSE;                         // 可用标志先清零 / Usable flag cleared first

(*------------------------------------------------------------------------------
 * 段 2｜非有限值防御：六个输入全查（含默认注入的大气压与新风比）
 *      Non-finite defense on all six inputs
 *-----------------------------------------------------------------------------*)
IF (fRaTempC <> fRaTempC) OR (ABS(fRaTempC) > DL_MIX_INF)
   OR (fRaHumRatio <> fRaHumRatio) OR (ABS(fRaHumRatio) > DL_MIX_INF)
   OR (fOaTempC <> fOaTempC) OR (ABS(fOaTempC) > DL_MIX_INF)
   OR (fOaHumRatio <> fOaHumRatio) OR (ABS(fOaHumRatio) > DL_MIX_INF)
   OR (fOaFrac <> fOaFrac) OR (ABS(fOaFrac) > DL_MIX_INF)
   OR (fPress <> fPress) OR (ABS(fPress) > DL_MIX_INF) THEN
    eErr   := 16#0002_3110;              // 故障级：输入非有限 / Fault: non-finite input
    bError := TRUE;                      // 置故障标志（R45 配对） / Raise the fault flag
    bValid := FALSE;                     // 输出不可用 / Outputs unusable
    RETURN;
END_IF

(*------------------------------------------------------------------------------
 * 段 3｜域外钳位：新风比 0~100、含湿量 >= 0，信息级共码 3101（R90）
 *      Out-of-domain clamping with a shared info code per R90
 *-----------------------------------------------------------------------------*)
IF (fOaFrac < DL_MIX_FRAC_MIN) OR (fOaFrac > DL_MIX_FRAC_MAX) THEN
    fFracEff := MIN(MAX(fOaFrac, DL_MIX_FRAC_MIN), DL_MIX_FRAC_MAX) / 100.0; // 新风比双侧钳位并转份额 / Two-sided fraction clamp, converted to share
    eErr := 16#0002_3101;                // 信息级：新风比已钳位（不置 bError） / Info: outdoor fraction clamped, no fault flag
ELSE
    fFracEff := fOaFrac / 100.0;         // 合法新风比转份额 [1] / Valid fraction converted to share [1]
END_IF
IF fRaHumRatio < 0.0 THEN
    fRaWEff := 0.0;                      // 回风含湿量负值钳 0（物理下界） / Negative return humidity ratio clamped to zero
    eErr := 16#0002_3101;                // 信息级：含湿量已钳位复用（R90） / Info: humidity ratio clamped, code reused
ELSE
    fRaWEff := fRaHumRatio;              // 合法回风含湿量原值生效 / Valid return humidity ratio applied as-is
END_IF
IF fOaHumRatio < 0.0 THEN
    fOaWEff := 0.0;                      // 新风含湿量负值钳 0（物理下界） / Negative outdoor humidity ratio clamped to zero
    eErr := 16#0002_3101;                // 信息级：含湿量已钳位复用（R90） / Info: humidity ratio clamped, code reused
ELSE
    fOaWEff := fOaHumRatio;              // 合法新风含湿量原值生效 / Valid outdoor humidity ratio applied as-is
END_IF

(*------------------------------------------------------------------------------
 * 段 4｜质量守恒加权主体：干球与含湿量分别按新风比加权
 *      Mass-conservation weighting for temperature and humidity ratio
 *-----------------------------------------------------------------------------*)
fMixTempC := fFracEff * fOaTempC + (1.0 - fFracEff) * fRaTempC; // 混合干球温度 [摄氏度] / Mixed dry-bulb temperature [degC]
fMixHumRatio := fFracEff * fOaWEff + (1.0 - fFracEff) * fRaWEff; // 混合含湿量 [kg 水蒸气/kg 干空气] / Mixed humidity ratio [kg/kg dry air]

(*------------------------------------------------------------------------------
 * 段 5｜混合焓内联复算（依赖收窄，见头注释段）：h = 1.006·T + W·(2501 + 1.86·T)
 *      Inline enthalpy per the dependency-narrowing declaration
 *-----------------------------------------------------------------------------*)
fMixEnthalpy := DL_MIX_CP_DRY * fMixTempC + fMixHumRatio * (DL_MIX_HFG0 + DL_MIX_CP_VAP * fMixTempC); // 混合比焓 [kJ/kg 干空气] / Mixed specific enthalpy [kJ/kg dry air]

(*------------------------------------------------------------------------------
 * 段 6｜结露判据：p_v_mix > p_ws(T_mix) 即越过饱和线（与 Magnus 反解温度
 *       比较法等价，免内联反解公式，饱和压取自族属主件）
 *       Condensation criterion via pressure comparison, owner FC sourced
 *-----------------------------------------------------------------------------*)
fDenom := DL_MIX_MW + fMixHumRatio;      // 分压反算分母 [kg/kg]，W >= 0 时恒 >= 0.622，仍强制闸 / Denominator, always >= 0.622 for W >= 0, still gated
IF fDenom <= DL_MIX_EPS THEN
    eErr   := 16#0002_3110;              // 故障级：分母退化复用非有限码（R90） / Fault: degenerate denominator, code reused
    bError := TRUE;                      // 置故障标志 / Raise the fault flag
    bValid := FALSE;                     // 输出不可用 / Outputs unusable
    RETURN;
END_IF
fPvMix := fMixHumRatio * fPress / fDenom; // 混合点水汽分压 [Pa] / Mixed vapor partial pressure [Pa]
IF (NOT FC_DL_VaporPressureSat(fTempC := fMixTempC, fPvSat => fPwsMix, bValid => _bPwsValid, bClamped => _bPwsClamped, eErr => _nPwsErr, bError => _bPwsError)) OR (NOT _bPwsValid) THEN
    eErr   := 16#0002_3110;              // 故障级：属主件拒绝复用（R90） / Fault: owner FC rejected, code reused
    bError := TRUE;                      // 置故障标志 / Raise the fault flag
    bValid := FALSE;                     // 输出不可用 / Outputs unusable
    RETURN;
END_IF
bCondensation := (fPvMix > fPwsMix);     // 结露预警（工况事实，不置故障） / Condensation warning, an operating fact, not a fault

bValid := TRUE;                          // 输出可用 / Outputs usable
FC_DL_MixAirStateCalc := TRUE;           // 返回 TRUE = 计算有效 / Return TRUE = computation valid
END_FUNCTION

(* ---- FC_DL_OvershootPctCalc.st ---- *)
// FC_DL_OvershootPctCalc v1.0.0
// 开源溯源：self-cleanroom / 回路 KPI 族
(*
  道莅工业代码库 | DL_Algo | FC_DL_OvershootPctCalc
  版本: 1.0.0 | 日期: 2026-11-23 | 轮次: R75
  功能: 阶跃响应超调量百分比：σ% = (y_peak − y_final)/(y_final − y_init) × 100；
        稳态幅差分母域闸；单调响应（无超调）返回负值按 0 收口
  邻件关系: 与 FC_DL_SettleTimeCalc（本批 S23，整定时间）成对 —— 差异点：
            超调件算峰值越界幅度，整定件算进入容差带时刻，两件共享
            阶跃响应特征入参口径（yInit/yFinal），码位独立
*)
FUNCTION FC_DL_OvershootPctCalc : REAL
VAR_INPUT
    fYInit    : REAL := 0.0;    // 阶跃前稳态值 [工程单位] / Pre-step steady value
    fYFinal   : REAL := 0.0;    // 目标稳态值 [工程单位] / Target steady value
    fYPeak    : REAL := 0.0;    // 响应峰值 [工程单位] / Response peak value
    fEps      : REAL := 1.0E-6; // 幅差判零容差 [工程单位] / Amplitude tolerance
END_VAR
VAR_OUTPUT
    bValid    : BOOL;           // 结果有效回执 [-] / Result validity receipt
    uErrorId  : UDINT;          // 事件码，0 = 无事件；16#0002_2901 = 域外/矛盾拒收 / Event code
END_VAR
VAR
    fDenom    : REAL;           // 分母 = y_final − y_init [工程单位] / Denominator
    fOver     : REAL;           // 超调绝对量 [工程单位] / Overshoot amount
    fResult   : REAL;           // 结果中间量 [%] / Result intermediate
END_VAR

// —— 段 0：全路径缺省 —— //
bValid := FALSE;                // 有效回执预清 / Validity preset
uErrorId := 16#0000;            // 事件码预清 / Event code preset
fOver := 0.0;                   // 超调量预清 / Overshoot preset
fResult := 0.0;                 // 结果预清 / Result preset
FC_DL_OvershootPctCalc := 0.0;  // 返回值缺省零 / Return default zero

// —— 段 1：非有限闸 —— //
IF (fYInit <> fYInit) OR (fYFinal <> fYFinal) OR (fYPeak <> fYPeak)
   OR (ABS(fYInit) >= 3.0E38) OR (ABS(fYFinal) >= 3.0E38) OR (ABS(fYPeak) >= 3.0E38) THEN
    uErrorId := 16#0002_2901;   // 输入非有限拒收 / Non-finite reject
    RETURN;
END_IF

// —— 段 2：分母域闸（R4：除法前判分母） —— //
fDenom := fYFinal - fYInit;     // 稳态幅差 [工程单位] / Steady amplitude difference
IF ABS(fDenom) < fEps THEN      // 幅差近零：阶跃幅值无效 / Near-zero step amplitude
    uErrorId := 16#0002_2901;   // 信息级：分母为零 / Info level: zero denominator
    RETURN;                     // 不计算返回 / Return without computation
END_IF

// —— 段 3：主计算（峰值须高于终值的正向超调口径） —— //
IF fDenom > 0.0 THEN
    fOver := fYPeak - fYFinal;  // 正向阶跃：峰值超终值量 / Positive step overshoot
ELSE
    fOver := fYFinal - fYPeak;  // 负向阶跃：口径镜像 / Negative step mirrored
END_IF
IF fOver <= 0.0 THEN
    fResult := 0.0;             // 无超调（单调响应）：按零收口 / No overshoot: zero
ELSE
    fResult := fOver / fDenom * 100.0;   // σ% = 超调量/幅差 ×100（分母非零已过闸）/ Overshoot percent
END_IF
FC_DL_OvershootPctCalc := fResult;   // 返回值 = 超调百分比 / Return equals overshoot percent
bValid := TRUE;                 // 有效回执 / Validity receipt
END_FUNCTION

(* ---- FC_DL_ParabolaVertexIterStep.st ---- *)
(* ============================================================
   DL_Algo / FC_DL_ParabolaVertexIterStep ｜ v1.0.0 ｜ 2026-11-25
   功能：抛物线插值顶点步。三点唯一确定抛物线，顶点横坐标
         xv = 0.5·[x1²(f2−f3)+x2²(f3−f1)+x3²(f1−f2)] / [x1(f2−f3)+x2(f3−f1)+x3(f1−f2)]；
         二阶系数 a（>0 为极小）由三点差商式给出，出 fCurv
   边界：横坐标重合（|Δx|≤1E-12）或分母近零（三点共线）→ bDegenerate=TRUE，
         fXv 取三点横坐标中位数、fCurv=0（N1：判据位与实值同源置位）
   依赖：仅 IEC 61131-3（ABS / MIN / MAX） ｜ 溯源：DLF-B-ROOTSTEP（内部原创线）
   ============================================================ *)
FUNCTION FC_DL_ParabolaVertexIterStep : BOOL
VAR_INPUT
    fX1 : LREAL;  // 第一点横坐标 [-] / Abscissa of the first point
    fX2 : LREAL;  // 第二点横坐标 [-] / Abscissa of the second point
    fX3 : LREAL;  // 第三点横坐标 [-] / Abscissa of the third point
    fF1 : LREAL;  // 第一点函数值 [-] / Function value of the first point
    fF2 : LREAL;  // 第二点函数值 [-] / Function value of the second point
    fF3 : LREAL;  // 第三点函数值 [-] / Function value of the third point
END_VAR
VAR_OUTPUT
    fXv         : LREAL;  // 顶点横坐标 [-] / Abscissa of the parabola vertex
    fCurv       : REAL;   // 二阶系数 a（>0 极小 / <0 极大）[-] / Quadratic coefficient
    bDegenerate : BOOL;   // 三点共线或横坐标重合 [-] / Collinear points or repeated abscissae
END_VAR
VAR
    _fNum  : LREAL;  // 顶点公式分子 [-] / Numerator of the vertex formula
    _fDen  : LREAL;  // 顶点公式分母 [-] / Denominator of the vertex formula
    _fDx12 : LREAL;  // x1 − x2 [-] / Difference of the first and second abscissae
    _fDx13 : LREAL;  // x1 − x3 [-] / Difference of the first and third abscissae
    _fDx23 : LREAL;  // x2 − x3 [-] / Difference of the second and third abscissae
    _fMid  : LREAL;  // 三点横坐标中位数 [-] / Median abscissa
END_VAR
VAR CONSTANT
    DL_PRV_EPS : LREAL := 1.0E-12;  // 分母判零容差 [-] / Denominator zero tolerance
END_VAR

(* 段 0：出口预置安全侧（顶点 0、曲率 0、标退化，N1/N3） *)
FC_DL_ParabolaVertexIterStep := FALSE;
fXv := 0.0;  fCurv := 0.0;  bDegenerate := TRUE;

(* 段 1：非有限闸（六个入参全量枚举） *)
IF (fX1 <> fX1) OR (fX2 <> fX2) OR (fX3 <> fX3)
   OR (fF1 <> fF1) OR (fF2 <> fF2) OR (fF3 <> fF3) THEN
    RETURN;
END_IF

(* 段 2：横坐标互异判据（三点必须互异） *)
_fDx12 := fX1 - fX2;  _fDx13 := fX1 - fX3;  _fDx23 := fX2 - fX3;
_fMid := MAX(MIN(fX1, fX2), MIN(MAX(fX1, fX2), fX3));   // 三数中位数
fXv := _fMid;                                          // 退化出口先落中位数
IF (ABS(_fDx12) <= DL_PRV_EPS) OR (ABS(_fDx13) <= DL_PRV_EPS) OR (ABS(_fDx23) <= DL_PRV_EPS) THEN
    RETURN;
END_IF

(* 段 3：顶点分子/分母与三点共线判据 *)
_fNum := fX1 * fX1 * (fF2 - fF3) + fX2 * fX2 * (fF3 - fF1) + fX3 * fX3 * (fF1 - fF2);
_fDen := fX1 * (fF2 - fF3) + fX2 * (fF3 - fF1) + fX3 * (fF1 - fF2);
IF ABS(_fDen) <= DL_PRV_EPS THEN RETURN; END_IF           // 共线：无唯一顶点

(* 段 4：顶点与二阶系数（除子已证非零） *)
fXv := 0.5 * _fNum / _fDen;
fCurv := LREAL_TO_REAL((fF1 * _fDx23 + fF2 * (fX3 - fX1) + fF3 * _fDx12)
        / (_fDx12 * _fDx13 * _fDx23));

(* 段 5：结果复检（判据位与实值同源，N4） *)
IF (fXv <> fXv) OR ((fXv - fXv) <> (fXv - fXv)) OR (fCurv <> fCurv) THEN
    fXv := _fMid;  fCurv := 0.0;  bDegenerate := TRUE;  RETURN;
END_IF
bDegenerate := FALSE;  FC_DL_ParabolaVertexIterStep := TRUE;
END_FUNCTION

(* ---- FC_DL_PidLambdaTune.st ---- *)
(*
  FC_DL_PidLambdaTune  —  IMC/λ 整定纯换算（FOPDT 三参数）/ IMC lambda tuning calculator
  分类 Category : DL_Algo
  码位 Code     : 16#02_3_83
  版本 Version  : 1.0.0
  来源 Source   : t2-1-lgf-math — IEC 61131-3 标准语义的道莅防御性实现
  溯源 Origin   : clean-room 实现，SIMC/IMC 公开整定公式，未复制任何源码行
                  （与 FB_DL_AutoTuneRelay 严格分工：本件只做纯换算不产生激励；在线辨识由 FB_DL_AutoTuneRelay 承载）
  功能 Function : 1) 由 FOPDT 三参数（K/T/τ）与闭环目标时间常数 λ 直接算 PID 系数：Kc = T/(K·(λ+τ))、Ti = MIN(T, 4·(λ+τ))；
                  2) 一阶对象默认不投微分（Td = 0）；bDerivativeOn 且 λ < τ 时按变体投 Td = τ/2；
                  3) 反向作用（K < 0）按 ABS(K) 计算并置信息码（符号语义由上层承接）；
                  4) 引脚命名对齐既有件 FB_DL_PidController（仅体例，不实例化）。
  边界 Boundary : ① fProcGain = 0 / fLambdaS <= 0 / fTimeConstS <= 0 / fDeadTimeS < 0 / fKcMax <= 0 均判组态错置码
                     且不输出系数（防除零与负增益误导，系数出口维持 0）；
                  ② λ < τ/2 判「整定过激」：bFeasible := FALSE 但仍给系数并置告警（是否采纳由工艺决定）；
                  ③ fKc 输出上限取 VAR_INPUT fKcMax（禁魔法数），越限钳制；
                  ④ K < 0 按 ABS(K) 计算并置「反向作用」信息码；
                  ⑤ 解除式自证：bFeasible 每调用重算，下一调用 λ 回到 >= τ/2 即自动解除（无锁存）；
                  ⑥ 本件为纯函数：无 VAR 记忆量、无定时器、无激励输出。
  依赖 Depends  : 仅 Standard.library（ABS/MIN）；引脚命名对齐 FB_DL_PidController（已注册）
  码表 Error codes（本件格 02_3_83，子码步进 +0x100）:
    16#0002_0183 信息级：反向作用（K < 0），已按 ABS(K) 计算
    16#0002_0283 故障级：组态非法（K = 0 / λ <= 0 / T <= 0 / τ < 0 / fKcMax <= 0），不输出系数
    16#0002_0383 告警级：λ < τ/2 整定过激（bFeasible = FALSE，系数仍给出）

  修订历史 Revision :
    2026-11-18  v1.0.0  R38 首版
*)

FUNCTION FC_DL_PidLambdaTune : BOOL
VAR_INPUT
    fProcGain    : REAL;              // 过程增益 K [无量纲]，域 <> 0 / Process gain, nonzero
    fTimeConstS  : REAL;              // 过程时间常数 T [s]，域 > 0 / Process time constant
    fDeadTimeS   : REAL;              // 纯滞后 τ [s]，域 >= 0 / Dead time
    fLambdaS     : REAL;              // 闭环目标时间常数 λ [s]，域 > 0 / Desired closed-loop time constant
    bDerivativeOn: BOOL := FALSE;     // 微分投用开关（λ < τ 时投 Td = τ/2 变体）/ Derivative enable variant
    fKcMax       : REAL;              // Kc 输出上限 [无量纲]，域 > 0（禁魔法数）/ Kc ceiling from configuration
END_VAR
VAR_OUTPUT
    fKc          : REAL;              // 比例增益 Kc [无量纲] / Proportional gain
    fTiS         : REAL;              // 积分时间 Ti [s] / Integral time
    fTdS         : REAL;              // 微分时间 Td [s] / Derivative time
    bFeasible    : BOOL;              // 整定可行标志（λ < τ/2 置 FALSE）/ Feasible flag
    nErrId       : UDINT;             // 事件码，0 = 无事件 / Event code, 0 = none
    fMsgCode     : REAL;              // 事件码 REAL 镜像（与 nErrId 同值，规格契约项）/ REAL mirror of the event code
END_VAR
VAR
    rKabs, rLam, rTau : LREAL;        // |K|/λ/τ 宽域暂存 / Wide-domain scratch of K, lambda, tau
    rSum              : LREAL;        // (λ + τ) 暂存 / Lambda plus tau
END_VAR

(* —— 段 1：输出缺省与组态闸（纯函数，每调用重算） —— *)
fKc := 0.0;  fTiS := 0.0;  fTdS := 0.0;    // 系数出口缺省 0（组态错不输出系数，规格强制）
bFeasible := TRUE;                          // 缺省可行
nErrId := 16#0000_0000;                     // 事件码缺省无事件
fMsgCode := 0.0;                            // REAL 镜像缺省 0
FC_DL_PidLambdaTune := FALSE;               // 返回值缺省失败

rKabs := LREAL(ABS(fProcGain));             // 按 |K| 计算（符号语义见段 4）
rLam  := LREAL(fLambdaS);
rTau  := LREAL(fDeadTimeS);

IF (rKabs < 1.0E-12) OR (rLam <= 0.0) OR (LREAL(fTimeConstS) <= 0.0)
   OR (rTau < 0.0) OR (LREAL(fKcMax) <= 0.0) THEN
    nErrId  := 16#0002_0283;                // 故障级：组态非法
    fMsgCode := 283.0;                      // REAL 镜像同步
    RETURN;                                 // 不输出系数（出口维持 0）
END_IF

(* —— 段 2：SIMC/λ 整定式（分母 rSum = λ + τ 已闸 > 0，无除零） —— *)
rSum := rLam + rTau;
fKc  := REAL(LREAL(fTimeConstS) / (rKabs * rSum));          // Kc = T / (|K|·(λ+τ))
fTiS := REAL(MIN(LREAL(fTimeConstS), 4.0 * rSum));          // Ti = MIN(T, 4·(λ+τ))
fTdS := 0.0;                                                // 一阶对象默认不投 D
IF bDerivativeOn AND (rLam < rTau) THEN
    fTdS := REAL(rTau / 2.0);                               // 微分变体：λ < τ 时投 Td = τ/2
END_IF

(* —— 段 3：Kc 上限钳制（上限来自 VAR_INPUT，禁魔法数） —— *)
IF LREAL(fKc) > LREAL(fKcMax) THEN
    fKc := fKcMax;                                          // 越上限钳制
END_IF

(* —— 段 4：符号与可行性判据（先信息码后告警码，互不覆盖故障） —— *)
IF fProcGain < 0.0 THEN
    nErrId := 16#0002_0183;                                 // 信息级：反向作用，已按 |K| 计算
END_IF
IF rLam < (rTau / 2.0) THEN
    bFeasible := FALSE;                                     // 整定过激：λ < τ/2
    nErrId := 16#0002_0383;                                 // 告警级：过激告警（系数仍给出，采纳由工艺决定）
END_IF

(* —— 段 5：出口与返回值 —— *)
fMsgCode := DINT_TO_REAL(DINT(nErrId));                     // REAL 镜像单点同步
FC_DL_PidLambdaTune := TRUE;                                // 换算已执行

END_FUNCTION

(* ---- FC_DL_PmvComfortIndex.st ---- *)
(*
  ==================================================================
  组件名 Component  : FC_DL_PmvComfortIndex
  分类   Category   : DL_Algo
  复杂度 Complexity  : 中
  版本   Version    : 1.0.1
  功能   Purpose    : PMV / PPD 热舒适指标计算（ISO 7730 公开 Fanger 六参数
                      公式链）。输入空气温度 / 平均辐射温度 / 空气流速 / 水
                      蒸汽分压 / 新陈代谢率 / 服装热阻，输出 PMV（钳 ±3）与
                      PPD（0..100%），供 HVAC 优化目标函数使用。
  来源   Source     : t1-oscat-building（热舒适域）
  溯源   Origin     : Fanger PMV 公式与 PPD 映射为 ISO 7730 公开标准公式链，
                      clean-room 自研实现，未复制 OSCAT 或任何厂商私有库
                      源码。
  平台   Platform   : 纯 IEC 61131-3，CODESYS / TwinCAT / InoProShop 通用
  分工声明 Split     : 与 FC_DL_HumidAirEnthalpy 分工——后者做湿空气焓值，本
                      件只做热舒适指标；与 FB_DL_NightPurgeSeq 分工——后者
                      为夜间吹扫顺控，本件为评价指标（无状态纯函数）。
  作者   Author     : 道莅代码库 · PLC 编程专家（R58）
  ------------------------------------------------------------------
  功能说明  : 四段式防御（R45）：预置 → 域闸门（六参数非有限 + ISO 7730 适用
              域：Ta/Tr 10..40 摄氏度，v 0..1 米每秒，pa 0..2.7 千帕，M 46.5..
              232 瓦每平方米，Icl 0..2 克罗，越域钳位信息级）→ 域内迭代求
              服装表面温度 tcl（固定 20 次迭代有界环，不动点收敛，无死循环
              风险）→ 结果非有限复检兜底。
  错误语义  : bError = TRUE 仅故障级（非有限入参）；bClamped = TRUE 信息级
              （六参数越域钳位，返回钳位口径结果）；bValid = TRUE 表示结果
              可用。
  修订记录  : 2026-11-21 v1.0.0 首次入库（R58 批 2 · 序号 6）
              2026-11-21 v1.0.1 R59 返修中①：段 6 补 fPpdPct 非有限/越界复检，拦负底数经 EXPT 的 NaN 穿透
*)
FUNCTION FC_DL_PmvComfortIndex : BOOL
VAR_INPUT
    fTaC   : LREAL; // 空气干球温度 [摄氏度]，域 10..40 / the air dry bulb temperature [degree celsius]
    fTrC   : LREAL; // 平均辐射温度 [摄氏度]，域 10..40 / the mean radiant temperature [degree celsius]
    fVaMs  : LREAL; // 空气流速 [米每秒]，域 0..1 / the air velocity [meter per second]
    fPaKpa : LREAL; // 水蒸汽分压 [千帕]，域 0..2.7 / the water vapour partial pressure [kilopascal]
    fMetW  : LREAL; // 新陈代谢率 [瓦每平方米]，域 46.5..232 / the metabolic rate [watt per square meter]
    fIclClo: LREAL; // 服装热阻 [克罗]，域 0..2 / the clothing insulation [clo]
END_VAR
VAR_OUTPUT
    fPmv    : LREAL; // PMV 预测平均投票（钳 ±3）[无量纲] / the predicted mean vote, clamped
    fPpdPct : LREAL; // PPD 预测不满意百分比 [百分数] / the predicted percentage dissatisfied [percent]
    bValid  : BOOL;  // 结果可用标志 [-] / the result usable flag
    bClamped: BOOL;  // 六参数越域钳位发生（信息级）[-] / an out of domain clamp happened, informational
    bError  : BOOL;  // 故障标志（非有限入参）[-] / the fault flag, a non finite input
END_VAR
VAR
    lrTa   : LREAL; // 空气温度工作量 [摄氏度] / the air temperature work value
    lrTr   : LREAL; // 辐射温度工作量 [摄氏度] / the radiant temperature work value
    lrVa   : LREAL; // 流速工作量 [米每秒] / the velocity work value
    lrPa   : LREAL; // 蒸汽分压工作量 [千帕] / the vapour pressure work value
    lrMet  : LREAL; // 新陈代谢工作量 [瓦每平方米] / the metabolic work value
    lrIcl  : LREAL; // 服装热阻工作量 [克罗] / the insulation work value
    lrMw   : LREAL; // 净机械功（本库取外部功为 0）[瓦每平方米] / the external work, zero in this library
    lrFcl  : LREAL; // 服装面积因子 [无量纲] / the clothing area factor
    lrTcl  : LREAL; // 服装表面温度迭代值 [摄氏度] / the clothing surface temperature iterate
    lrTclN : LREAL; // 服装表面温度下一迭代值 [摄氏度] / the next clothing surface iterate
    lrHc   : LREAL; // 对流换热系数 [瓦每平方米每开尔文] / the convective heat transfer coefficient
    lrLoad : LREAL; // 热负荷项 [瓦每平方米] / the thermal load term
    lrPmvW : LREAL; // PMV 未钳工作量 [无量纲] / the unclamped PMV work value
    nI     : DINT;  // 固定迭代索引 [次] / the fixed iteration index
END_VAR
VAR CONSTANT
    DL_PMV_ITER   : DINT  := 20;                 // 服装温度定点迭代次数 [次]（有界环，无死循环）/ the clothing temperature fixed iterations
    DL_PMV_RELAX  : LREAL := 0.75;               // 迭代松弛因子 [无量纲]，防定点振荡 / the iteration relaxation factor
    DL_PMV_ABSMAX : LREAL := 3.0;                // PMV 出口钳位界 [无量纲] / the PMV clamp bound
    DL_PMV_TAMIN  : LREAL := 10.0;               // 空气温度域下界 [摄氏度] / the air temperature floor
    DL_PMV_TAMAX  : LREAL := 40.0;               // 空气温度域上界 [摄氏度] / the air temperature ceiling
    DL_PMV_VAMAX  : LREAL := 1.0;                // 流速域上界 [米每秒] / the velocity ceiling
    DL_PMV_PAMAX  : LREAL := 2.7;                // 蒸汽分压域上界 [千帕] / the vapour pressure ceiling
    DL_PMV_METMIN : LREAL := 46.5;               // 新陈代谢域下界 [瓦每平方米] / the metabolic floor
    DL_PMV_METMAX : LREAL := 232.0;              // 新陈代谢域上界 [瓦每平方米] / the metabolic ceiling
    DL_PMV_ICLMAX : LREAL := 2.0;                // 服装热阻域上界 [克罗] / the insulation ceiling
END_VAR

// 段 1｜返回值与错误状态预置安全值（四段式第一段，R45）/ segment 1, preset the return and error states
FC_DL_PmvComfortIndex := FALSE; // 受理标志预置假 / preset the accepted flag false
fPmv := 0.0; // PMV 预置中性零 / preset the PMV neutral zero
fPpdPct := 5.0; // PPD 预置下限 5%（PMV = 0 的对应值）/ preset the PPD floor five percent
bValid := FALSE; // 有效标志预置假 / preset the valid flag false
bClamped := FALSE; // 钳位标志预置假 / preset the clamp flag false
bError := FALSE; // 故障标志预置假 / preset the fault flag false

// 段 2｜非有限入参闸（六参数自反双判据全覆盖，R79 / R151）/ segment 2, the non finite gate over the six inputs
IF (fTaC <> fTaC) OR ((fTaC - fTaC) <> (fTaC - fTaC)) THEN // 空气温度非有限 / a non finite air temperature
    bError := TRUE; // 置故障标志（R45 配对）/ raise the fault flag
END_IF
IF (fTrC <> fTrC) OR ((fTrC - fTrC) <> (fTrC - fTrC)) THEN // 辐射温度非有限 / a non finite radiant temperature
    bError := TRUE; // 置故障标志 / raise the fault flag
END_IF
IF (fVaMs <> fVaMs) OR ((fVaMs - fVaMs) <> (fVaMs - fVaMs)) THEN // 流速非有限 / a non finite velocity
    bError := TRUE; // 置故障标志 / raise the fault flag
END_IF
IF (fPaKpa <> fPaKpa) OR ((fPaKpa - fPaKpa) <> (fPaKpa - fPaKpa)) THEN // 蒸汽分压非有限 / a non finite vapour pressure
    bError := TRUE; // 置故障标志 / raise the fault flag
END_IF
IF (fMetW <> fMetW) OR ((fMetW - fMetW) <> (fMetW - fMetW)) THEN // 新陈代谢非有限 / a non finite metabolic rate
    bError := TRUE; // 置故障标志 / raise the fault flag
END_IF
IF (fIclClo <> fIclClo) OR ((fIclClo - fIclClo) <> (fIclClo - fIclClo)) THEN // 服装热阻非有限 / a non finite insulation
    bError := TRUE; // 置故障标志 / raise the fault flag
END_IF
IF bError THEN // 非有限命中：返回预置安全值 / a non finite hit, return the preset safe values
    RETURN; // 早退 / return early
END_IF

// 段 3｜ISO 7730 适用域钳位（信息级，越域判据按方向分列 R146）/ segment 3, the applicability clamps, informational
lrTa := fTaC; // 装空气温度 / load the air temperature
IF lrTa < DL_PMV_TAMIN THEN // 低于下界 / below the floor
    lrTa := DL_PMV_TAMIN; // 钳到下界 / clamp to the floor
    bClamped := TRUE; // 信息级钳位 / the informational clamp
ELSIF lrTa > DL_PMV_TAMAX THEN // 高于上界 / above the ceiling
    lrTa := DL_PMV_TAMAX; // 钳到上界 / clamp to the ceiling
    bClamped := TRUE; // 信息级钳位 / the informational clamp
END_IF
lrTr := fTrC; // 装辐射温度 / load the radiant temperature
IF lrTr < DL_PMV_TAMIN THEN // 低于下界 / below the floor
    lrTr := DL_PMV_TAMIN; // 钳到下界 / clamp to the floor
    bClamped := TRUE; // 信息级钳位 / the informational clamp
ELSIF lrTr > DL_PMV_TAMAX THEN // 高于上界 / above the ceiling
    lrTr := DL_PMV_TAMAX; // 钳到上界 / clamp to the ceiling
    bClamped := TRUE; // 信息级钳位 / the informational clamp
END_IF
lrVa := fVaMs; // 装流速 / load the velocity
IF lrVa < 0.0 THEN // 负流速（物理不可达，钳零）/ a negative velocity, clamped to zero
    lrVa := 0.0; // 钳到零 / clamp to zero
    bClamped := TRUE; // 信息级钳位 / the informational clamp
ELSIF lrVa > DL_PMV_VAMAX THEN // 高于上界 / above the ceiling
    lrVa := DL_PMV_VAMAX; // 钳到上界 / clamp to the ceiling
    bClamped := TRUE; // 信息级钳位 / the informational clamp
END_IF
lrPa := fPaKpa; // 装蒸汽分压 / load the vapour pressure
IF lrPa < 0.0 THEN // 负分压钳零 / a negative pressure clamped to zero
    lrPa := 0.0; // 钳到零 / clamp to zero
    bClamped := TRUE; // 信息级钳位 / the informational clamp
ELSIF lrPa > DL_PMV_PAMAX THEN // 高于上界 / above the ceiling
    lrPa := DL_PMV_PAMAX; // 钳到上界 / clamp to the ceiling
    bClamped := TRUE; // 信息级钳位 / the informational clamp
END_IF
lrMet := fMetW; // 装新陈代谢率 / load the metabolic rate
IF lrMet < DL_PMV_METMIN THEN // 低于下界 / below the floor
    lrMet := DL_PMV_METMIN; // 钳到下界 / clamp to the floor
    bClamped := TRUE; // 信息级钳位 / the informational clamp
ELSIF lrMet > DL_PMV_METMAX THEN // 高于上界 / above the ceiling
    lrMet := DL_PMV_METMAX; // 钳到上界 / clamp to the ceiling
    bClamped := TRUE; // 信息级钳位 / the informational clamp
END_IF
lrIcl := fIclClo; // 装服装热阻 / load the insulation
IF lrIcl < 0.0 THEN // 负热阻钳零 / a negative insulation clamped to zero
    lrIcl := 0.0; // 钳到零 / clamp to zero
    bClamped := TRUE; // 信息级钳位 / the informational clamp
ELSIF lrIcl > DL_PMV_ICLMAX THEN // 高于上界 / above the ceiling
    lrIcl := DL_PMV_ICLMAX; // 钳到上界 / clamp to the ceiling
    bClamped := TRUE; // 信息级钳位 / the informational clamp
END_IF

// 段 4｜服装面积因子与服装表面温度定点迭代（固定 20 次有界环）/ segment 4, the area factor and the clothing temperature iteration
IF lrIcl <= 0.5 THEN // 低热阻面积因子分支（ISO 7730 公开分段）/ the low insulation branch
    lrFcl := 1.0 + 0.2 * lrIcl; // 面积因子 / the area factor
ELSE // 高热阻面积因子分支 / the high insulation branch
    lrFcl := 1.05 + 0.1 * lrIcl; // 面积因子 / the area factor
END_IF
lrTcl := lrTa; // 迭代初值取空气温度（安全侧收敛起点）/ the iterate starts at the air temperature
lrMw := 0.0; // 本库外部机械功取零（坐立轻活动场景）/ the external work is zero in this library
FOR nI := 1 TO DL_PMV_ITER DO // 固定界迭代环，无死循环风险 / the fixed bound iteration loop
    lrHc := 12.1 * SQRT(lrVa); // 对流换热候选一（流速项）/ the convective candidate one
    IF 2.38 * EXPT(ABS(lrTcl - lrTa), 0.25) > lrHc THEN // 候选二更大则取大（ISO 7730 取大规则）/ take the larger candidate
        lrHc := 2.38 * EXPT(ABS(lrTcl - lrTa), 0.25); // 取候选二 / take the candidate two
    END_IF
    lrTclN := 35.7 - 0.028 * (lrMet - lrMw) - 0.155 * lrIcl * (3.96E-8 * lrFcl * (EXPT(lrTcl + 273.15, 4.0) - EXPT(lrTr + 273.15, 4.0)) + lrFcl * lrHc * (lrTcl - lrTa)); // ISO 7730 标准隐式定点式（右端含 tcl，靠固定环迭代收敛）/ the ISO 7730 implicit fixed point form, converged by the fixed loop
    lrTcl := lrTcl + DL_PMV_RELAX * (lrTclN - lrTcl); // 松弛更新 / the relaxed update
END_FOR

// 段 5｜PMV 主式与 PPD 映射（ISO 7730 公开公式链）/ segment 5, the PMV formula and the PPD mapping
lrHc := 12.1 * SQRT(lrVa); // 出口段对流系数重算（与迭代末值口径一致）/ the outlet convective coefficient
IF 2.38 * EXPT(ABS(lrTcl - lrTa), 0.25) > lrHc THEN // 取大规则 / the larger rule
    lrHc := 2.38 * EXPT(ABS(lrTcl - lrTa), 0.25); // 取候选二 / take the candidate two
END_IF
lrLoad := (lrMet - lrMw) // 热负荷项组装（Fanger 展开式）/ assemble the thermal load
        - 3.05E-3 * (5733.0 - 6.99 * (lrMet - lrMw) - lrPa * 1000.0) // 呼吸显热项（分压换算帕）/ the respiration sensible term
        - 0.42 * ((lrMet - lrMw) - 58.15) // 呼吸潜热项 / the respiration latent term
        - 1.7E-5 * lrMet * (5867.0 - lrPa * 1000.0) // 皮肤蒸发项 / the skin evaporation term
        - 0.0014 * lrMet * (34.0 - lrTa) // 皮肤对流项 / the skin convection term
        - 3.96E-8 * lrFcl * (EXPT(lrTcl + 273.15, 4.0) - EXPT(lrTr + 273.15, 4.0)) // 辐射项 / the radiation term
        - lrFcl * lrHc * (lrTcl - lrTa); // 服装对流项 / the clothing convection term
lrPmvW := (0.303 * EXP(-0.036 * lrMet) + 0.028) * lrLoad; // PMV 权重式 / the PMV weighted form
IF lrPmvW > DL_PMV_ABSMAX THEN // PMV 上钳 / clamp the PMV up
    fPmv := DL_PMV_ABSMAX; // 钳到上界 / clamp to the bound
ELSIF lrPmvW < -DL_PMV_ABSMAX THEN // PMV 下钳 / clamp the PMV down
    fPmv := -DL_PMV_ABSMAX; // 钳到下界 / clamp to the bound
ELSE // 域内直通 / inside the domain
    fPmv := lrPmvW; // 直通结果 / pass through
END_IF
fPpdPct := 100.0 - 95.0 * EXP(-0.03353 * EXPT(fPmv, 4.0) - 0.2179 * fPmv * fPmv); // PPD 映射式 / the PPD mapping

// 段 6｜结果非有限复检兜底（防御纵深，正常路径不可达）/ segment 6, the result recheck as defense in depth
IF (fPmv <> fPmv) OR ((fPmv - fPmv) <> (fPmv - fPmv)) THEN // PMV 非有限 / a non finite PMV
    fPmv := 0.0; // 归中性零 / zero to the neutral
    fPpdPct := 5.0; // PPD 回下限 / the PPD to the floor
    bValid := FALSE; // 降有效标志 / drop the valid flag
    RETURN; // 早退（受理标志保持假）/ return early, refused
END_IF
// R59 修 R58 中①：fPpdPct 复检三件套（负底数经 EXPT(fPmv,4.0) 可产生 NaN 穿透，PMV 复检不覆盖本输出）
IF (fPpdPct <> fPpdPct) OR ((fPpdPct - fPpdPct) <> (fPpdPct - fPpdPct)) THEN // PPD 非有限（NOT ISFINITE 等价自反判式）/ a non finite PPD
    fPpdPct := 5.0; // 回安全下限 / to the safe floor
    bValid := FALSE; // 降有效标志 / drop the valid flag
    RETURN; // 早退（受理标志保持假）/ return early, refused
END_IF
IF fPpdPct < 0.0 THEN // 负 PPD 钳零（信息级）/ a negative PPD clamped to zero
    fPpdPct := 0.0; bClamped := TRUE; // 钳到下界 0 并置信息级 / clamp to the floor zero
ELSIF fPpdPct > 100.0 THEN // 越上界回夹到 [0,100] / above the ceiling, re-clamped into the band
    fPpdPct := 100.0; bClamped := TRUE; // 钳到上界 100 并置信息级 / clamp to the ceiling hundred
END_IF
bValid := TRUE; // 结果可用 / the result usable
FC_DL_PmvComfortIndex := TRUE; // 求解受理 / accept the result
END_FUNCTION

(* ---- FC_DL_PolishPadPressureCalc.st ---- *)
(*
  DL Factory R88 | FC_DL_PolishPadPressureCalc
  功能：算抛光垫比压 p=F/A，A=πD²/4，N/mm² 按 ×1000 换算 kPa，并按 5~30 kPa 判带宽
  开源溯源：无（clean-room 自研，依据公开工艺公式 圆盘接触比压式 p=F/(πD²/4)，许可证=MIT，借鉴点=公式结构）
  规则：R1-R16 全遵守；R88 简单件标量形（纯标量入参出参，无循环体、无方法、无属性、无数组）
*)
FUNCTION FC_DL_PolishPadPressureCalc : REAL
VAR_INPUT
    fForceN : REAL := 300.0; // 抛光下压力 F [N] / polishing down force [N]
    fDiaMm : REAL := 200.0; // 抛光垫（或工件）接触直径 D [mm] / pad or workpiece diameter [mm]
    fMinKPa : REAL := 5.0; // 比压允许下限（工艺带宽） [kPa] / lower pressure band [kPa]
    fMaxKPa : REAL := 30.0; // 比压允许上限（工艺带宽） [kPa] / upper pressure band [kPa]
END_VAR
VAR_OUTPUT
    fPressKPa : REAL; // 抛光垫比压 p [kPa] / pad specific pressure [kPa]
    xInBand : BOOL; // TRUE=比压落在允许带宽内 [-] / TRUE when inside the band [-]
END_VAR
VAR
    fAreaMm2 : REAL; // 接触面积 A=πD²/4（除零判据） [mm²] / contact area, the divisor [mm^2]
    fPressMpa : REAL; // 比压 N/mm²（数值等同 MPa） [N/mm²] / specific pressure [N/mm^2]
END_VAR

// 段 1｜出口预置
FC_DL_PolishPadPressureCalc := -1.0; // 哨兵返回 -1（无效） [-] / sentinel return -1, invalid [-]
fPressKPa := 0.0; // 比压预置零 [kPa] / pressure preset zero [kPa]
xInBand := FALSE; // 带宽位预置 FALSE [-] / band flag preset false [-]
fAreaMm2 := 0.0; // 接触面积预置零 [mm²] / area preset zero [mm^2]
fPressMpa := 0.0; // 比压中间量预置零 [N/mm²] / pressure mid value preset zero [N/mm^2]

// 段 2｜非有限拦截 + 域闸
IF NOT (fForceN > -1.0E30 AND fForceN < 1.0E30) OR NOT (fDiaMm > -1.0E30 AND fDiaMm < 1.0E30) THEN
    RETURN; // 下压力/直径任一非有限即拒算 [-] / any non finite input rejected [-]
END_IF
IF NOT (fMinKPa > -1.0E30 AND fMinKPa < 1.0E30) OR NOT (fMaxKPa > -1.0E30 AND fMaxKPa < 1.0E30) THEN
    RETURN; // 带宽上下限任一非有限则判据静默失效，故先拦 [kPa] / band limits must be finite [kPa]
END_IF
IF fForceN < 0.0 OR fDiaMm < 1.0E-9 THEN
    RETURN; // 力非负闸 + 直径正域闸（面积分母不得为零） [N, mm] / non negative force and positive diameter
END_IF
IF fMinKPa <= 0.0 OR fMaxKPa <= fMinKPa THEN
    RETURN; // 带宽自洽闸：下限须为正、上限须严格大于下限 [kPa] / band consistency gate [kPa]
END_IF

// 段 3｜计算
fAreaMm2 := 3.14159265 * fDiaMm * fDiaMm * 0.25; // 无量纲 × mm² × 0.25 = mm²，A=πD²/4（乘 0.25 替除 4） [mm²] / [mm^2]
IF fAreaMm2 < 1.0E-9 THEN
    RETURN; // 除法前分母闸：面积必须大于 1E-9 才可作除数 [mm²] / denominator gate before the division [mm^2]
END_IF
fPressMpa := fForceN / fAreaMm2; // N ÷ mm² = N/mm²（数值等同 MPa） [N/mm²] / [N] / [mm^2] = [N/mm^2]
fPressKPa := fPressMpa * 1000.0; // N/mm² × 1000 = kPa（1 N/mm²=1 MPa=1000 kPa） [kPa] / [kPa]

// 段 4｜判定与饱和
IF NOT (fPressKPa > -1.0E30 AND fPressKPa < 1.0E30) THEN
    RETURN; // 结果非有限再拦一次 [-] / re-check the result for finiteness [-]
END_IF
xInBand := (fPressKPa >= fMinKPa) AND (fPressKPa <= fMaxKPa); // 双侧闭区间直比 [kPa] / closed two sided band compare [kPa]

// 段 5｜出口自检
IF fPressKPa < 0.0 THEN
    RETURN; // 出口自检：比压不得为负（负值说明力符号错） [kPa] / pressure must not be negative [kPa]
END_IF
FC_DL_PolishPadPressureCalc := fPressKPa; // 返回抛光垫比压 [kPa] / return the pad specific pressure [kPa]
END_FUNCTION

(* ---- FC_DL_RegulaFalsiIterStep.st ---- *)
(* ============================================================
   DL_Algo / FC_DL_RegulaFalsiIterStep ｜ v1.0.0 ｜ 2026-11-25
   功能：试位法（弦线法）单步：x = fA − fFa·(fB−fA)/(fFb−fFa) 并夹回括号；
         同时出「新点入括号后保守宽度上界」MAX(x−a, b−x)（本件不求值 f(x)）
   边界：差分 < fDenEps（含入参≤0 时取内部下限）或两端同号 → 退二分中点；
         任一入参非有限 → 新点写 0、宽度 0（N1：实值与判据同拍改写）
   依赖：仅 IEC 61131-3（ABS / MIN / MAX / LIMIT） ｜ 溯源：DLF-B-ROOTSTEP（内部原创线）
   ============================================================ *)
FUNCTION FC_DL_RegulaFalsiIterStep : BOOL
VAR_INPUT
    fA      : LREAL;  // 括号下界 [-] / Lower bracket bound
    fB      : LREAL;  // 括号上界 [-] / Upper bracket bound
    fFa     : LREAL;  // 下界函数值 [-] / Function value at the lower bound
    fFb     : LREAL;  // 上界函数值 [-] / Function value at the upper bound
    fDenEps : LREAL;  // 差分下限（防零），建议 > 0 [-] / Minimum difference guarding the division
END_VAR
VAR_OUTPUT
    fXnew     : LREAL;  // 弦线插值新点（已夹回括号）[-] / Interpolated point clamped into the bracket
    fWidthNew : LREAL;  // 保守宽度上界 [-] / Conservative width upper bound
END_VAR
VAR
    _fDen  : LREAL;  // 弦线分母 = fFb − fFa [-] / Chord slope denominator
    _fEps  : LREAL;  // 生效判零下限 [-] / Effective denominator floor
    _fLo   : LREAL;  // 括号小端 [-] / Smaller bracket end
    _fHi   : LREAL;  // 括号大端 [-] / Larger bracket end
    _fMid  : LREAL;  // 二分中点 [-] / Bisection midpoint
END_VAR
VAR CONSTANT
    DL_RGZ_FLOOR : LREAL := 1.0E-12;  // 差分判零内部下限 [-] / Internal floor for the denominator
END_VAR

(* 段 0：出口预置安全侧（新点 0、宽度 0，防 NaN 直穿） *)
FC_DL_RegulaFalsiIterStep := FALSE;
fXnew := 0.0;  fWidthNew := 0.0;

(* 段 1：非有限闸（原始入参判定） *)
IF (fA <> fA) OR (fB <> fB) OR (fFa <> fFa) OR (fFb <> fFb) OR (fDenEps <> fDenEps) THEN
    RETURN;
END_IF
IF ((fB - fA) - (fB - fA)) <> ((fB - fA) - (fB - fA)) THEN RETURN; END_IF

(* 段 2：括号排序、中点与退化处理 *)
_fLo := MIN(fA, fB);  _fHi := MAX(fA, fB);
_fMid := _fLo + (_fHi - _fLo) / 2.0;
fXnew := _fMid;                               // 缺省即二分中点
IF (_fHi - _fLo) <= DL_RGZ_FLOOR THEN RETURN; END_IF

(* 段 3：分母与括号有效性（不可解均退二分，不置错） *)
IF fDenEps > DL_RGZ_FLOOR THEN _fEps := fDenEps; ELSE _fEps := DL_RGZ_FLOOR; END_IF
_fDen := fFb - fFa;
IF ABS(_fDen) <= _fEps THEN
    fWidthNew := MAX(_fMid - _fLo, _fHi - _fMid);
    FC_DL_RegulaFalsiIterStep := TRUE;  RETURN;
END_IF
IF ((fFa > 0.0) AND (fFb > 0.0)) OR ((fFa < 0.0) AND (fFb < 0.0)) THEN
    fWidthNew := MAX(_fMid - _fLo, _fHi - _fMid);   // 同号：括号失效，退二分
    FC_DL_RegulaFalsiIterStep := TRUE;  RETURN;
END_IF

(* 段 4：弦线插值并夹回括号（夹界即 N4 出口闸），除子已证 |den| > _fEps *)
fXnew := LIMIT(_fLo, fA - fFa * (fB - fA) / _fDen, _fHi);
fWidthNew := MAX(fXnew - _fLo, _fHi - fXnew);

(* 段 5：结果复检 *)
IF (fXnew <> fXnew) OR ((fXnew - fXnew) <> (fXnew - fXnew)) THEN
    fXnew := _fMid;  fWidthNew := 0.0;  RETURN;
END_IF
FC_DL_RegulaFalsiIterStep := TRUE;
END_FUNCTION

(* ---- FC_DL_RhFromDewPoint.st ---- *)
//==============================================================================
// 函数：FC_DL_RhFromDewPoint ｜ 中文名称：露点→相对湿度逆运算原子（焓湿图族拆分④）
// 所属子库：DL_Algo ｜ 版本：v1.0.1 ｜ 兼容：CODESYS V3.5+ / TwinCAT 3 / 汇川 InoProShop
// 功能描述：RH = 100·p_ws(Td)/p_ws(T)，纯比值运算；两次调用族属主
//           FC_DL_VaporPressureSat，本件无自带公式常量（零内联公式）。
//           与 FC_DL_DewPointCalc 构成双向对，round-trip 验收向量：
//           DewPoint→Rh→DewPoint 误差 < 1E-3 °C。
// 开源溯源 (Origin)：改写自 OSCAT Building 行为定义（OSCAT 许可，仅行为定义，零代码行）——道莅 clean-room 实现
// 单位表：T[°C] / Td[°C] / RH[%] / p_ws[Pa]
// 错误码表：16#0002_3001 信息级（露点超干球钳 100 或干球温度已钳位，不置
//           bError）/ 16#0002_3010 故障级（露点超干球 > 5 K 传感器矛盾或
//           输入非有限，置 bError）/ 16#0002_3002、16#0002_3011、
//           16#0002_3012 预留禁用（不得挪用）
// 状态机：N/A（纯函数，无状态）
// 边界行为：① Td 略超 T（<= 5 K）→ 过饱和物理矛盾按饱和处理：RH 钳 100 +
//           信息 3001，不置故障（比值语义可安全钳位——与
//           FC_DL_HumidityRatioCalc 的 2E11 故障策略差异：该件分母直接
//           参与除法必须故障保护，本件纯比值无发散风险）；② Td 超干球
//           5 K 以上判传感器矛盾 → 故障 3010、bValid := FALSE；③ 输入
//           非有限 → 故障 3010 复用（R90）；④ 干球温度域外（−40~100 °C
//           外）→ 钳位 + 信息 3001 复用（R90）；⑤ 属主件拒绝 → 故障 3010
//           复用；异常路径输出确定值 0，绝不输出未初始化值。
// 修订历史：v1.0.0 2026-11-17 首版（R23 派单 · T1-2 焓湿图族拆分④ · 双向对闭环）
//           v1.0.1 2026-11-23 R73 补 bValid 回执：段 5 两处属主件调用补收
//           bValid 局部回执，回执无效并入既有 3010 兜底分支，契约不变。
//==============================================================================

(*------------------------------------------------------------------------------
 * 调用示例：bOk := FC_DL_RhFromDewPoint(fTempC := 25.0, fDewPointC := 16.7,
 *                                       fRh => fRhPct, eErr => uE);
 * round-trip 验收：FC_DL_DewPointCalc(T, Rh) 得 Td 后经本件反解，RH 复现
 * 误差 < 1E-3 百分数；误差超限说明两件口径漂移，应停用并查常量属主。
 *-----------------------------------------------------------------------------*)
FUNCTION FC_DL_RhFromDewPoint : BOOL
VAR_INPUT
    fTempC     : LREAL;                  // 干球温度 [摄氏度]，有效域 -40.0..100.0，域外钳位照算 / Dry-bulb temperature [degC], valid range -40.0..100.0
    fDewPointC : LREAL;                  // 露点温度 [摄氏度] / Dew-point temperature [degC]
END_VAR
VAR_OUTPUT
    fRh        : LREAL;                  // 相对湿度 [百分数]，输出域 0..100 / Relative humidity [percent], output range 0..100
    eErr       : UDINT;                  // 错误码，0 = 无错 / Error code, 0 = no error
    bError     : BOOL;                   // 故障级标志，仅故障级错误置位 / Fault-class flag, set only on fault-level codes
    bValid     : BOOL;                   // 输出可用标志 / Outputs usable flag
END_VAR
VAR CONSTANT
    DL_RHDP_TMIN     : LREAL := -40.0;   // 干球温度钳位下限 [摄氏度]，对齐族属主有效域 / Dry-bulb clamp floor [degC], aligned with the family owner domain
    DL_RHDP_TMAX     : LREAL := 100.0;   // 干球温度钳位上限 [摄氏度] / Dry-bulb clamp ceiling [degC]
    DL_RHDP_OVERHYST : LREAL := 5.0;     // 传感器矛盾判据阈 [摄氏度]，露点超干球此值即故障 / Sensor contradiction threshold [degC]
    DL_RHDP_INF      : LREAL := 1.7976931348623157E308; // LREAL 幅值上限 / LREAL magnitude ceiling
END_VAR
VAR
    fTEff    : LREAL;                    // 钳位后的生效干球温度 [摄氏度] / Effective clamped dry-bulb temperature [degC]
    fPwsDb   : LREAL;                    // 干球温度下饱和压 [Pa] / Saturation pressure at the dry bulb [Pa]
    fPwsTd   : LREAL;                    // 露点温度下饱和压 [Pa] / Saturation pressure at the dew point [Pa]
    _bPwsValid : BOOL;                   // 饱和压属主件输出可用回执 / Saturation owner FC outputs-usable receipt
    _bPwsClamped : BOOL;    // 属主件钳位回执（本件不消费，仅契约全回执） / Owner clamp receipt (unused, full-receipt contract)
    _nPwsErr     : UDINT;   // 属主件错误码回执 / Owner error-code receipt
    _bPwsError   : BOOL;    // 属主件故障级回执 / Owner fault-flag receipt
END_VAR

(*------------------------------------------------------------------------------
 * 段 1｜出口默认值：入口即赋确定值
 *      Exit defaults: outputs assigned deterministically on entry
 *-----------------------------------------------------------------------------*)
FC_DL_RhFromDewPoint := FALSE;           // 返回值默认无效 / Return value preset invalid
fRh := 0.0;                              // 相对湿度默认置零 / Relative humidity preset to zero
eErr := 16#0000_0000;                    // 错误码先清零 / Error code cleared first
bError := FALSE;                         // 故障标志先清零 / Fault flag cleared first
bValid := FALSE;                         // 可用标志先清零 / Usable flag cleared first

(*------------------------------------------------------------------------------
 * 段 2｜非有限值防御（NaN 用 (x<>x)，Inf 用双侧幅值判，R79）
 *      Non-finite defense per R79
 *-----------------------------------------------------------------------------*)
IF (fTempC <> fTempC) OR (ABS(fTempC) > DL_RHDP_INF)
   OR (fDewPointC <> fDewPointC) OR (ABS(fDewPointC) > DL_RHDP_INF) THEN
    eErr   := 16#0002_3010;              // 故障级：输入非有限复用传感器矛盾码（R90） / Fault: non-finite input, code reused
    bError := TRUE;                      // 置故障标志（R45 配对） / Raise the fault flag
    bValid := FALSE;                     // 输出不可用 / Outputs unusable
    RETURN;
END_IF

(*------------------------------------------------------------------------------
 * 段 3｜干球温度钳位：域外信息级照算（R90 复用 3001）
 *      Dry-bulb clamping, info code reused per R90
 *-----------------------------------------------------------------------------*)
IF (fTempC < DL_RHDP_TMIN) OR (fTempC > DL_RHDP_TMAX) THEN
    fTEff := MIN(MAX(fTempC, DL_RHDP_TMIN), DL_RHDP_TMAX); // 双侧钳位到有效域 / Two-sided clamp into valid range
    eErr := 16#0002_3001;                // 信息级：温度已钳位（不置 bError） / Info: temperature clamped, no fault flag
ELSE
    fTEff := fTempC;                     // 合法温度原值生效 / Valid temperature applied as-is
END_IF

(*------------------------------------------------------------------------------
 * 段 4｜传感器矛盾闸：Td 超干球 5 K 以上 → 故障；略超（<= 5 K）→ 钳 100
 *      先判重故障再判轻矛盾，两级策略次序不可反
 *      Sensor contradiction gate, severe case checked before the mild one
 *-----------------------------------------------------------------------------*)
IF fDewPointC > (fTEff + DL_RHDP_OVERHYST) THEN
    fRh := 0.0;                          // 矛盾输入丢弃，输出确定值 0 / Contradictory input discarded, output zero
    eErr   := 16#0002_3010;              // 故障级：露点超干球 > 5 K，判传感器矛盾 / Fault: dew point exceeds dry bulb by more than 5 K
    bError := TRUE;                      // 置故障标志 / Raise the fault flag
    bValid := FALSE;                     // 输出不可用 / Outputs unusable
    RETURN;
ELSIF fDewPointC > fTEff THEN
    fRh := 100.0;                        // 过饱和物理矛盾按饱和处理（比值语义安全钳位） / Supersaturation treated as saturation, safe ratio clamp
    IF eErr = 16#0000_0000 THEN
        eErr := 16#0002_3001;            // 信息级：露点超干球钳 100（不置 bError） / Info: dew point above dry bulb, clamped to 100
    END_IF
    bValid := TRUE;                      // 输出可用（钳位结论可用） / Outputs usable
    FC_DL_RhFromDewPoint := TRUE;        // 返回 TRUE = 计算有效 / Return TRUE = computation valid
    RETURN;
END_IF

(*------------------------------------------------------------------------------
 * 段 5｜双向对主体：RH = 100·p_ws(Td)/p_ws(T)，两次调用族属主件
 *      Round-trip core via two owner FC calls, denominator guarded
 *-----------------------------------------------------------------------------*)
IF (NOT FC_DL_VaporPressureSat(fTempC := fTEff, fPvSat => fPwsDb, bValid => _bPwsValid, bClamped => _bPwsClamped, eErr => _nPwsErr, bError => _bPwsError)) OR (NOT _bPwsValid) THEN
    eErr   := 16#0002_3010;              // 故障级：属主件拒绝复用（R90） / Fault: owner FC rejected, code reused
    bError := TRUE;                      // 置故障标志 / Raise the fault flag
    bValid := FALSE;                     // 输出不可用 / Outputs unusable
    RETURN;
END_IF
IF (NOT FC_DL_VaporPressureSat(fTempC := fDewPointC, fPvSat => fPwsTd, bValid => _bPwsValid, bClamped => _bPwsClamped, eErr => _nPwsErr, bError => _bPwsError)) OR (NOT _bPwsValid) THEN
    eErr   := 16#0002_3010;              // 故障级：属主件拒绝复用（R90） / Fault: owner FC rejected, code reused
    bError := TRUE;                      // 置故障标志 / Raise the fault flag
    bValid := FALSE;                     // 输出不可用 / Outputs unusable
    RETURN;
END_IF
IF ABS(fPwsDb) <= 1.0E-6 THEN
    eErr   := 16#0002_3010;              // 故障级：分母退化复用（域内理论上恒正，仍强制闸） / Fault: degenerate denominator, guarded even if theoretically positive
    bError := TRUE;                      // 置故障标志 / Raise the fault flag
    bValid := FALSE;                     // 输出不可用 / Outputs unusable
    RETURN;
END_IF
fRh := 100.0 * fPwsTd / fPwsDb;          // 相对湿度 [百分数] / Relative humidity [percent]
IF fRh > 100.0 THEN
    fRh := 100.0;                        // 数值越界钳回 100（浮点噪声防护） / Numerical overshoot clamped to 100
END_IF
IF fRh < 0.0 THEN
    fRh := 0.0;                          // 数值越界钳回 0（浮点噪声防护） / Numerical undershoot clamped to 0
END_IF
bValid := TRUE;                          // 输出可用 / Outputs usable
FC_DL_RhFromDewPoint := TRUE;            // 返回 TRUE = 计算有效 / Return TRUE = computation valid
END_FUNCTION

(* ---- FC_DL_ScannerReadRateCalc.st ---- *)
(*
  DL Factory R83 | FC_DL_ScannerReadRateCalc
  功能：按读码总次数与首读成功数算首读率，并算失败件平均重读次数与未读率。
  开源溯源：无（clean-room 自研，依据公开工艺公式，来源=行业通用公式，许可证=MIT，借鉴点=公式结构）
  规则：R1-R21 全遵守
*)
FUNCTION FC_DL_ScannerReadRateCalc : REAL
VAR_INPUT
    diTotal   : DINT; // 读码总次数（含重读）[次] / Total read attempts incl. retries [-]
    diFirstOk : DINT; // 首次即读成功次数 [次] / First-attempt successes [-]
    diRetry   : DINT; // 重读累计次数 [次] / Total retries [-]
    diNoRead  : DINT; // 最终未读次数 [次] / Final no-reads [-]
END_VAR
VAR_OUTPUT
    fFsrPct    : REAL; // 首读率 FSR [%] / First-scan rate [%]
    fAvgRetry  : REAL; // 失败件平均重读次数 [次/件] / Mean retries per failed read [-]
    fNoReadPct : REAL; // 最终未读率 [%] / Final no-read rate [%]
    xValid     : BOOL; // 计算有效性标志 / Calculation validity flag
END_VAR
VAR
    diFail : DINT; // 首读失败件数 [次] / First-read failures [-]
END_VAR
// 出口预置：四出口统一预置（R256）
fFsrPct := 0.0; fAvgRetry := 0.0; fNoReadPct := 0.0; xValid := FALSE;
// 计数器域闸：任一项为负或首读超总数即判采集异常（整数无 NaN，仍做符号与次序检查）
IF diTotal <= 0 OR diFirstOk < 0 OR diRetry < 0 OR diNoRead < 0 OR diFirstOk > diTotal OR diNoRead > diTotal THEN
    FC_DL_ScannerReadRateCalc := -1.0; RETURN;  // 哨兵 -1：计数域越界 / Sentinel -1: counter domain violation
END_IF
// 首读率：首读成功 ÷ 总次数 × 100（先转 REAL 再除，避免整数截断）
fFsrPct := (DINT_TO_REAL(diFirstOk) / DINT_TO_REAL(diTotal)) * 100.0; // 首读率 [%] / First-scan rate
// 首读失败件数：总数 - 首读成功，非负由上面的次序闸保证
diFail := diTotal - diFirstOk;     // 首读失败数 [次] / First-read failures [-]
// 平均重读：重读次数 ÷ 失败件数，分母分支显式判零（R4/R21）
IF diFail > 0 THEN                 // 失败件数分母显式零闸 / Explicit zero gate on failure count
    fAvgRetry := DINT_TO_REAL(diRetry) / DINT_TO_REAL(diFail); // 平均重读 [次/件] / Mean retries
ELSE
    fAvgRetry := 0.0;               // 全首读通过，无重读 / All first-read, no retries
END_IF
// 未读率：未读次数 ÷ 总次数 × 100（总次数已判正）
fNoReadPct := (DINT_TO_REAL(diNoRead) / DINT_TO_REAL(diTotal)) * 100.0; // 未读率 [%] / No-read rate
xValid := TRUE;                           // 链路有效 / Chain valid
FC_DL_ScannerReadRateCalc := fFsrPct;     // 返回首读率 [%] / Return first-scan rate [%]
END_FUNCTION

(* ---- FC_DL_SCurveTimeOptCalc.st ---- *)
(*
  Name: FC_DL_SCurveTimeOptCalc
  Category: DL_Algo
  Version: 1.0.0
  Round: R89 / 2026-11-25
  开源溯源：clean-room 自研（族 运动规划算法，ST 开源生态实测 0 命中，无外部代码引入）
  功能：S 曲线七段最短时间规划（速度/加速度/加加速度三重约束），含距离不足时降速（三角速度）分支与退化处置。
  边界条件：① 三入参全部过非有限闸；速度/加速度/加加速度任一 ≤ 0 判组态非法，返回哨兵 -1（时间不可表）；
            ② 距离 ≤ 1E-9 mm 视为零行程：时间/峰值/两时长为 0、段数 0、xValid = TRUE、xDistTooShort = TRUE；
            ③ 七段可达判据：2×加速段距离 ≤ 行程 时存在匀速段（段数 7）；否则对峰值速度做 40 次二分求根，
               峰值速度收敛到 1E-6 相对精度以内（禁 EXPT 原语：拐点平方根已用 SQRT 展开，R140 委托纪律）；
            ④ 段数口径：7 = 加加速/恒加速/减加速 + 匀速 + 加减速/恒减速/减减速；6 = 无匀速且恒加速段非零；
               4 = 无匀速且恒加速段为零（三角加速）；三者互斥完备；
            ⑤ 全部钳位/饱和仅作用于量值（时长、段数），有效性由 xValid 单独表达，不伪造事实。
  量纲自证：mm/s² ÷ mm/s³ = s；mm/s ÷ mm/s² = s；mm/s × s = mm；距离[m] ÷ 速度[m/s] = s。
*)
FUNCTION FC_DL_SCurveTimeOptCalc : REAL
VAR_INPUT
    fDistMm : REAL;         (* 行程 [mm] Travel distance [mm] *)
    fVmaxMmS : REAL;        (* 速度上限 [mm/s] Velocity limit [mm/s] *)
    fAmaxMmS2 : REAL;       (* 加速度上限 [mm/s2] Acceleration limit [mm/s2] *)
    fJmaxMmS3 : REAL;       (* 加加速度上限 [mm/s3] Jerk limit [mm/s3] *)
END_VAR
VAR_OUTPUT
    fTimeS : REAL;          (* 最短时间 [s] Minimum time [s] *)
    fVpeakMmS : REAL;       (* 规划峰值速度 [mm/s] Planned peak velocity [mm/s] *)
    fTjS : REAL;            (* 加加速（jerk）段时长 [s] Jerk phase duration [s] *)
    fTaS : REAL;            (* 恒加速段时长（0 = 无） [s] Constant acceleration duration [s] *)
    nSegCount : INT;        (* 段数（0/4/6/7） [段] Segment count *)
    xValid : BOOL;          (* 计算有效性标志 [-] Calculation valid flag *)
    xDistTooShort : BOOL;   (* 距离不足以达到速度上限（已降速） [-] Velocity limit not reachable *)
END_VAR
VAR CONSTANT
    DL_SCV_EPS : REAL := 1.0E-9;        (* 判据容差 [-] Criterion tolerance *)
    DL_SCV_ITER : INT := 40;            (* 二分迭代次数（相对精度 < 1E-6） [次] Bisection iterations *)
    DL_SCV_HALF : REAL := 2.0;          (* 对称行程除数 [-] Symmetric travel divisor *)
    DL_SCV_ZNUM : INT := 0;             (* 零段数 [-] Zero segment count *)
    DL_SCV_N4 : INT := 4;               (* 四段（三角加速、无匀速） [段] Four segments *)
    DL_SCV_N6 : INT := 6;               (* 六段（恒加速段非零、无匀速） [段] Six segments *)
    DL_SCV_N7 : INT := 7;               (* 七段（含匀速段） [段] Seven segments *)
END_VAR
VAR
    fVlim : REAL := 0.0;    (* 达恒加速度所需速度（A²/J） [mm/s] Velocity to reach Amax [mm/s] *)
    fTj : REAL := 0.0;      (* 加加速段时长 [s] Jerk phase duration [s] *)
    fTa : REAL := 0.0;      (* 恒加速段时长 [s] Constant acceleration duration [s] *)
    fTv : REAL := 0.0;      (* 匀速段时长 [s] Constant velocity duration [s] *)
    fDacc : REAL := 0.0;    (* 单个加速段距离 [mm] Single acceleration distance [mm] *)
    fVpeak : REAL := 0.0;   (* 峰值速度 [mm/s] Peak velocity [mm/s] *)
    fVlo : REAL := 0.0;     (* 二分下界 [mm/s] Bisection lower bound [mm/s] *)
    fVhi : REAL := 0.0;     (* 二分上界 [mm/s] Bisection upper bound [mm/s] *)
    fVmid : REAL := 0.0;    (* 二分中点 [mm/s] Bisection midpoint [mm/s] *)
    fTjC : REAL := 0.0;     (* 候选加加速时长 [s] Candidate jerk duration [s] *)
    fTaC : REAL := 0.0;     (* 候选恒加速时长 [s] Candidate accel duration [s] *)
    fDmid : REAL := 0.0;    (* 候选中点对应加速距离 [mm] Candidate accel distance [mm] *)
    nIter : INT := 1;       (* 二分迭代计数 [-] Bisection counter *)
END_VAR
(* 出口预置：七出口统一预置（R256） *)
fTimeS := 0.0; fVpeakMmS := 0.0; fTjS := 0.0; fTaS := 0.0;
nSegCount := DL_SCV_ZNUM; xValid := FALSE; xDistTooShort := FALSE;
(* 非有限闸：NaN 自反判 + Inf 差值自减判，三入参全枚举 *)
IF (fDistMm <> fDistMm) OR ((fDistMm - fDistMm) <> 0.0)
   OR (fVmaxMmS <> fVmaxMmS) OR ((fVmaxMmS - fVmaxMmS) <> 0.0)
   OR (fAmaxMmS2 <> fAmaxMmS2) OR ((fAmaxMmS2 - fAmaxMmS2) <> 0.0)
   OR (fJmaxMmS3 <> fJmaxMmS3) OR ((fJmaxMmS3 - fJmaxMmS3) <> 0.0) THEN
    FC_DL_SCurveTimeOptCalc := -1.0;         (* 哨兵 -1：入参非有限 / Sentinel -1, non-finite input *)
    RETURN;
END_IF
(* 组态域闸：三重上限任一为 0 即退化（时间不可表），距离不得为负 *)
IF (fVmaxMmS <= DL_SCV_EPS) OR (fAmaxMmS2 <= DL_SCV_EPS) OR (fJmaxMmS3 <= DL_SCV_EPS)
   OR (fDistMm < 0.0) THEN
    FC_DL_SCurveTimeOptCalc := -1.0;         (* 哨兵 -1：三重上限退化 / Sentinel -1, degenerate limits *)
    RETURN;
END_IF
(* 零行程退化：全部输出 0，段数 0，有效性置真（零距离是合法事实，不是错误） *)
IF fDistMm <= DL_SCV_EPS THEN
    xValid := TRUE;
    xDistTooShort := TRUE;
    nSegCount := DL_SCV_ZNUM;
    FC_DL_SCurveTimeOptCalc := 0.0;
    RETURN;
END_IF
(* 达恒加速度所需速度：A²/J，量纲 mm/s *)
fVlim := (fAmaxMmS2 * fAmaxMmS2) / fJmaxMmS3;
(* 先试速度上限 V：算其加速段距离，判断是否存在匀速段 *)
IF fVmaxMmS >= fVlim THEN
    fTj := fAmaxMmS2 / fJmaxMmS3;                       (* s = (mm/s2)/(mm/s3) *)
    fTa := (fVmaxMmS / fAmaxMmS2) - fTj;                (* 恒加速段，量纲 s *)
    fDacc := fVmaxMmS * ((DL_SCV_HALF * fTj) + fTa) / DL_SCV_HALF;   (* mm/s × s = mm *)
ELSE
    fTj := SQRT(fVmaxMmS / fJmaxMmS3);                  (* 三角加速：v = J·tj² *)
    fTa := 0.0;
    fDacc := fVmaxMmS * fTj;
END_IF
IF (DL_SCV_HALF * fDacc) <= fDistMm THEN
    fVpeak := fVmaxMmS;                                 (* 速度上限可达 / Limit reachable *)
ELSE
    (* 距离不足：对峰值速度二分求根，使 2×加速段距离 = 行程（单调增，故二分收敛） *)
    fVlo := 0.0;
    fVhi := fVmaxMmS;
    FOR nIter := 1 TO DL_SCV_ITER DO
        fVmid := (fVlo + fVhi) / DL_SCV_HALF;
        IF fVmid >= fVlim THEN
            fTjC := fAmaxMmS2 / fJmaxMmS3;
            fTaC := (fVmid / fAmaxMmS2) - fTjC;
            fDmid := fVmid * ((DL_SCV_HALF * fTjC) + fTaC) / DL_SCV_HALF;
        ELSE
            fTjC := SQRT(fVmid / fJmaxMmS3);
            fTaC := 0.0;
            fDmid := fVmid * fTjC;
        END_IF
        IF (DL_SCV_HALF * fDmid) > fDistMm THEN
            fVhi := fVmid;                              (* 距离超了：峰值取小 / Too far, lower bound *)
        ELSE
            fVlo := fVmid;                              (* 距离不足：峰值取大 / Too short, raise bound *)
        END_IF
    END_FOR
    fVpeak := fVlo;                                     (* 取保守下界，保证不超行程 / Conservative bound *)
END_IF
(* 按最终峰值速度复算 tj / ta / 单段加速距离 *)
IF fVpeak >= fVlim THEN
    fTj := fAmaxMmS2 / fJmaxMmS3;
    fTa := (fVpeak / fAmaxMmS2) - fTj;
    fDacc := fVpeak * ((DL_SCV_HALF * fTj) + fTa) / DL_SCV_HALF;
ELSE
    fTj := SQRT(fVpeak / fJmaxMmS3);
    fTa := 0.0;
    fDacc := fVpeak * fTj;
END_IF
(* 匀速段：剩余行程 ÷ 峰值速度（峰值已过正性闸，绝无零除） *)
IF fVpeak <= DL_SCV_EPS THEN
    FC_DL_SCurveTimeOptCalc := -1.0;         (* 哨兵 -1：峰值速度塌零（行程过小无法表出） / Degenerate *)
    RETURN;
END_IF
fTv := (fDistMm - (DL_SCV_HALF * fDacc)) / fVpeak;
IF fTv < 0.0 THEN
    fTv := 0.0;                                         (* 二分残差导致的微负归零 / Residual to zero *)
END_IF
(* 总时间：2×(加加速 + 恒加速 + 加加速) + 匀速 = 2×(2·tj+ta) + tv，量纲 s *)
fTimeS := DL_SCV_HALF * ((DL_SCV_HALF * fTj) + fTa) + fTv;
(* 段数判定：匀速段 > 0 → 7；否则看恒加速段是否为零 → 6 或 4 *)
IF fTv > DL_SCV_EPS THEN
    nSegCount := DL_SCV_N7;
ELSIF fTa > DL_SCV_EPS THEN
    nSegCount := DL_SCV_N6;
ELSE
    nSegCount := DL_SCV_N4;
END_IF
fVpeakMmS := fVpeak;
fTjS := fTj;
fTaS := fTa;
xDistTooShort := fVpeak < (fVmaxMmS - DL_SCV_EPS);
xValid := TRUE;                                        (* 链路有效 / Chain valid *)
FC_DL_SCurveTimeOptCalc := fTimeS;
END_FUNCTION
